(* IEC 61131-3 sources: IEC61131-3_ST_SCL_Mutation_Generator/Tests/mutatedCodeTraffic (part 2) *)

(* ---- M133.st ---- *)
FUNCTION_BLOCK TRAFFIC_CTRL

VAR_INPUT
    PedestrianButton1 : BOOL;
    PedestrianButton2 : BOOL;
END_VAR

VAR_OUTPUT
    NorthSouthRed : BOOL;
    NorthSouthYellow : BOOL;
    NorthSouthGreen : BOOL;
    EastWestRed : BOOL;
    EastWestYellow : BOOL;
    EastWestGreen : BOOL;
    PedestrianLight1 : BOOL;
    PedestrianLight2 : BOOL;
END_VAR

VAR
    LightState : INT := 0; (* 0: North-South Green, 1: North-South Yellow, 2: East-West Green, 3: East-West Yellow *)
    PedestrianRequest1 : BOOL := FALSE;
    PedestrianRequest2 : BOOL := FALSE;
    PedestrianCrossing : BOOL := FALSE;
    Timer : TON;
END_VAR

(* Check for pedestrian requests *)
IF PedestrianButton1 THEN
    PedestrianRequest1 := TRUE;
END_IF;

IF PedestrianButton2 THEN
    PedestrianRequest2 := TRUE;
END_IF;

(* Traffic light state machine *)
CASE LightState OF
    0: (* North-South Green *)
        NorthSouthGreen := TRUE;
        EastWestRed := TRUE;
        IF PedestrianRequest1 OR PedestrianRequest2 THEN
            Timer(IN := TRUE, PT := T#2s); (* Pedestrian crossing grace period *)
            IF Timer.Q THEN
                Timer(IN := FALSE);
                LightState := 2; (* MUTATED: CONST_VALUE_REPLACE *)
            END_IF;
        END_IF;

    1: (* North-South Yellow *)
        NorthSouthYellow := TRUE;
        EastWestRed := TRUE;
        Timer(IN := TRUE, PT := T#2s); (* Yellow light duration *)
        IF Timer.Q THEN
            Timer(IN := FALSE);
            LightState := 2;
        END_IF;

    2: (* East-West Green *)
        EastWestGreen := TRUE;
        NorthSouthRed := TRUE;
        IF PedestrianRequest1 THEN
            PedestrianLight1 := TRUE;
            PedestrianCrossing := TRUE;
        END_IF;
        IF PedestrianRequest2 THEN
            PedestrianLight2 := TRUE;
            PedestrianCrossing := TRUE;
        END_IF;
        IF PedestrianCrossing THEN
            Timer(IN := TRUE, PT := T#2s); (* Pedestrian crossing period *)
            IF Timer.Q THEN
                Timer(IN := FALSE);
                PedestrianRequest1 := FALSE;
                PedestrianRequest2 := FALSE;
                PedestrianLight1 := FALSE;
                PedestrianLight2 := FALSE;
                PedestrianCrossing := FALSE;
                LightState := 3;
            END_IF;
        END_IF;

    3: (* East-West Yellow *)
        EastWestYellow := TRUE;
        NorthSouthRed := TRUE;
        Timer(IN := TRUE, PT := T#2s); (* Yellow light duration *)
        IF Timer.Q THEN
            Timer(IN := FALSE);
            LightState := 0;
        END_IF;

END_CASE;

END_FUNCTION_BLOCK

(* ---- M134.st ---- *)
FUNCTION_BLOCK TRAFFIC_CTRL

VAR_INPUT
    PedestrianButton1 : BOOL;
    PedestrianButton2 : BOOL;
END_VAR

VAR_OUTPUT
    NorthSouthRed : BOOL;
    NorthSouthYellow : BOOL;
    NorthSouthGreen : BOOL;
    EastWestRed : BOOL;
    EastWestYellow : BOOL;
    EastWestGreen : BOOL;
    PedestrianLight1 : BOOL;
    PedestrianLight2 : BOOL;
END_VAR

VAR
    LightState : INT := 0; (* 0: North-South Green, 1: North-South Yellow, 2: East-West Green, 3: East-West Yellow *)
    PedestrianRequest1 : BOOL := FALSE;
    PedestrianRequest2 : BOOL := FALSE;
    PedestrianCrossing : BOOL := FALSE;
    Timer : TON;
END_VAR

(* Check for pedestrian requests *)
IF PedestrianButton1 THEN
    PedestrianRequest1 := TRUE;
END_IF;

IF PedestrianButton2 THEN
    PedestrianRequest2 := TRUE;
END_IF;

(* Traffic light state machine *)
CASE LightState OF
    0: (* North-South Green *)
        NorthSouthGreen := TRUE;
        EastWestRed := TRUE;
        IF PedestrianRequest1 OR PedestrianRequest2 THEN
            Timer(IN := TRUE, PT := T#2s); (* Pedestrian crossing grace period *)
            IF Timer.Q THEN
                Timer(IN := FALSE);
                LightState := 1;
            END_IF;
        END_IF;

    2: (* North-South Yellow *) (* MUTATED: CONST_VALUE_REPLACE *)
        NorthSouthYellow := TRUE;
        EastWestRed := TRUE;
        Timer(IN := TRUE, PT := T#2s); (* Yellow light duration *)
        IF Timer.Q THEN
            Timer(IN := FALSE);
            LightState := 2;
        END_IF;

    2: (* East-West Green *)
        EastWestGreen := TRUE;
        NorthSouthRed := TRUE;
        IF PedestrianRequest1 THEN
            PedestrianLight1 := TRUE;
            PedestrianCrossing := TRUE;
        END_IF;
        IF PedestrianRequest2 THEN
            PedestrianLight2 := TRUE;
            PedestrianCrossing := TRUE;
        END_IF;
        IF PedestrianCrossing THEN
            Timer(IN := TRUE, PT := T#2s); (* Pedestrian crossing period *)
            IF Timer.Q THEN
                Timer(IN := FALSE);
                PedestrianRequest1 := FALSE;
                PedestrianRequest2 := FALSE;
                PedestrianLight1 := FALSE;
                PedestrianLight2 := FALSE;
                PedestrianCrossing := FALSE;
                LightState := 3;
            END_IF;
        END_IF;

    3: (* East-West Yellow *)
        EastWestYellow := TRUE;
        NorthSouthRed := TRUE;
        Timer(IN := TRUE, PT := T#2s); (* Yellow light duration *)
        IF Timer.Q THEN
            Timer(IN := FALSE);
            LightState := 0;
        END_IF;

END_CASE;

END_FUNCTION_BLOCK

(* ---- M135.st ---- *)
FUNCTION_BLOCK TRAFFIC_CTRL

VAR_INPUT
    PedestrianButton1 : BOOL;
    PedestrianButton2 : BOOL;
END_VAR

VAR_OUTPUT
    NorthSouthRed : BOOL;
    NorthSouthYellow : BOOL;
    NorthSouthGreen : BOOL;
    EastWestRed : BOOL;
    EastWestYellow : BOOL;
    EastWestGreen : BOOL;
    PedestrianLight1 : BOOL;
    PedestrianLight2 : BOOL;
END_VAR

VAR
    LightState : INT := 0; (* 0: North-South Green, 1: North-South Yellow, 2: East-West Green, 3: East-West Yellow *)
    PedestrianRequest1 : BOOL := FALSE;
    PedestrianRequest2 : BOOL := FALSE;
    PedestrianCrossing : BOOL := FALSE;
    Timer : TON;
END_VAR

(* Check for pedestrian requests *)
IF PedestrianButton1 THEN
    PedestrianRequest1 := TRUE;
END_IF;

IF PedestrianButton2 THEN
    PedestrianRequest2 := TRUE;
END_IF;

(* Traffic light state machine *)
CASE LightState OF
    0: (* North-South Green *)
        NorthSouthGreen := TRUE;
        EastWestRed := TRUE;
        IF PedestrianRequest1 OR PedestrianRequest2 THEN
            Timer(IN := TRUE, PT := T#2s); (* Pedestrian crossing grace period *)
            IF Timer.Q THEN
                Timer(IN := FALSE);
                LightState := 1;
            END_IF;
        END_IF;

    1: (* North-South Yellow *)
        NorthSouthYellow := TRUE;
        EastWestRed := TRUE;
        Timer(IN := TRUE, PT := T#2s); (* Yellow light duration *)
        IF Timer.Q THEN
            Timer(IN := FALSE);
            LightState := 3; (* MUTATED: CONST_VALUE_REPLACE *)
        END_IF;

    2: (* East-West Green *)
        EastWestGreen := TRUE;
        NorthSouthRed := TRUE;
        IF PedestrianRequest1 THEN
            PedestrianLight1 := TRUE;
            PedestrianCrossing := TRUE;
        END_IF;
        IF PedestrianRequest2 THEN
            PedestrianLight2 := TRUE;
            PedestrianCrossing := TRUE;
        END_IF;
        IF PedestrianCrossing THEN
            Timer(IN := TRUE, PT := T#2s); (* Pedestrian crossing period *)
            IF Timer.Q THEN
                Timer(IN := FALSE);
                PedestrianRequest1 := FALSE;
                PedestrianRequest2 := FALSE;
                PedestrianLight1 := FALSE;
                PedestrianLight2 := FALSE;
                PedestrianCrossing := FALSE;
                LightState := 3;
            END_IF;
        END_IF;

    3: (* East-West Yellow *)
        EastWestYellow := TRUE;
        NorthSouthRed := TRUE;
        Timer(IN := TRUE, PT := T#2s); (* Yellow light duration *)
        IF Timer.Q THEN
            Timer(IN := FALSE);
            LightState := 0;
        END_IF;

END_CASE;

END_FUNCTION_BLOCK

(* ---- M136.st ---- *)
FUNCTION_BLOCK TRAFFIC_CTRL

VAR_INPUT
    PedestrianButton1 : BOOL;
    PedestrianButton2 : BOOL;
END_VAR

VAR_OUTPUT
    NorthSouthRed : BOOL;
    NorthSouthYellow : BOOL;
    NorthSouthGreen : BOOL;
    EastWestRed : BOOL;
    EastWestYellow : BOOL;
    EastWestGreen : BOOL;
    PedestrianLight1 : BOOL;
    PedestrianLight2 : BOOL;
END_VAR

VAR
    LightState : INT := 0; (* 0: North-South Green, 1: North-South Yellow, 2: East-West Green, 3: East-West Yellow *)
    PedestrianRequest1 : BOOL := FALSE;
    PedestrianRequest2 : BOOL := FALSE;
    PedestrianCrossing : BOOL := FALSE;
    Timer : TON;
END_VAR

(* Check for pedestrian requests *)
IF PedestrianButton1 THEN
    PedestrianRequest1 := TRUE;
END_IF;

IF PedestrianButton2 THEN
    PedestrianRequest2 := TRUE;
END_IF;

(* Traffic light state machine *)
CASE LightState OF
    0: (* North-South Green *)
        NorthSouthGreen := TRUE;
        EastWestRed := TRUE;
        IF PedestrianRequest1 OR PedestrianRequest2 THEN
            Timer(IN := TRUE, PT := T#2s); (* Pedestrian crossing grace period *)
            IF Timer.Q THEN
                Timer(IN := FALSE);
                LightState := 1;
            END_IF;
        END_IF;

    1: (* North-South Yellow *)
        NorthSouthYellow := TRUE;
        EastWestRed := TRUE;
        Timer(IN := TRUE, PT := T#2s); (* Yellow light duration *)
        IF Timer.Q THEN
            Timer(IN := FALSE);
            LightState := 2;
        END_IF;

    3: (* East-West Green *) (* MUTATED: CONST_VALUE_REPLACE *)
        EastWestGreen := TRUE;
        NorthSouthRed := TRUE;
        IF PedestrianRequest1 THEN
            PedestrianLight1 := TRUE;
            PedestrianCrossing := TRUE;
        END_IF;
        IF PedestrianRequest2 THEN
            PedestrianLight2 := TRUE;
            PedestrianCrossing := TRUE;
        END_IF;
        IF PedestrianCrossing THEN
            Timer(IN := TRUE, PT := T#2s); (* Pedestrian crossing period *)
            IF Timer.Q THEN
                Timer(IN := FALSE);
                PedestrianRequest1 := FALSE;
                PedestrianRequest2 := FALSE;
                PedestrianLight1 := FALSE;
                PedestrianLight2 := FALSE;
                PedestrianCrossing := FALSE;
                LightState := 3;
            END_IF;
        END_IF;

    3: (* East-West Yellow *)
        EastWestYellow := TRUE;
        NorthSouthRed := TRUE;
        Timer(IN := TRUE, PT := T#2s); (* Yellow light duration *)
        IF Timer.Q THEN
            Timer(IN := FALSE);
            LightState := 0;
        END_IF;

END_CASE;

END_FUNCTION_BLOCK

(* ---- M137.st ---- *)
FUNCTION_BLOCK TRAFFIC_CTRL

VAR_INPUT
    PedestrianButton1 : BOOL;
    PedestrianButton2 : BOOL;
END_VAR

VAR_OUTPUT
    NorthSouthRed : BOOL;
    NorthSouthYellow : BOOL;
    NorthSouthGreen : BOOL;
    EastWestRed : BOOL;
    EastWestYellow : BOOL;
    EastWestGreen : BOOL;
    PedestrianLight1 : BOOL;
    PedestrianLight2 : BOOL;
END_VAR

VAR
    LightState : INT := 0; (* 0: North-South Green, 1: North-South Yellow, 2: East-West Green, 3: East-West Yellow *)
    PedestrianRequest1 : BOOL := FALSE;
    PedestrianRequest2 : BOOL := FALSE;
    PedestrianCrossing : BOOL := FALSE;
    Timer : TON;
END_VAR

(* Check for pedestrian requests *)
IF PedestrianButton1 THEN
    PedestrianRequest1 := TRUE;
END_IF;

IF PedestrianButton2 THEN
    PedestrianRequest2 := TRUE;
END_IF;

(* Traffic light state machine *)
CASE LightState OF
    0: (* North-South Green *)
        NorthSouthGreen := TRUE;
        EastWestRed := TRUE;
        IF PedestrianRequest1 OR PedestrianRequest2 THEN
            Timer(IN := TRUE, PT := T#2s); (* Pedestrian crossing grace period *)
            IF Timer.Q THEN
                Timer(IN := FALSE);
                LightState := 1;
            END_IF;
        END_IF;

    1: (* North-South Yellow *)
        NorthSouthYellow := TRUE;
        EastWestRed := TRUE;
        Timer(IN := TRUE, PT := T#2s); (* Yellow light duration *)
        IF Timer.Q THEN
            Timer(IN := FALSE);
            LightState := 2;
        END_IF;

    2: (* East-West Green *)
        EastWestGreen := TRUE;
        NorthSouthRed := TRUE;
        IF PedestrianRequest1 THEN
            PedestrianLight1 := TRUE;
            PedestrianCrossing := TRUE;
        END_IF;
        IF PedestrianRequest2 THEN
            PedestrianLight2 := TRUE;
            PedestrianCrossing := TRUE;
        END_IF;
        IF PedestrianCrossing THEN
            Timer(IN := TRUE, PT := T#2s); (* Pedestrian crossing period *)
            IF Timer.Q THEN
                Timer(IN := FALSE);
                PedestrianRequest1 := FALSE;
                PedestrianRequest2 := FALSE;
                PedestrianLight1 := FALSE;
                PedestrianLight2 := FALSE;
                PedestrianCrossing := FALSE;
                LightState := 4; (* MUTATED: CONST_VALUE_REPLACE *)
            END_IF;
        END_IF;

    3: (* East-West Yellow *)
        EastWestYellow := TRUE;
        NorthSouthRed := TRUE;
        Timer(IN := TRUE, PT := T#2s); (* Yellow light duration *)
        IF Timer.Q THEN
            Timer(IN := FALSE);
            LightState := 0;
        END_IF;

END_CASE;

END_FUNCTION_BLOCK

(* ---- M138.st ---- *)
FUNCTION_BLOCK TRAFFIC_CTRL

VAR_INPUT
    PedestrianButton1 : BOOL;
    PedestrianButton2 : BOOL;
END_VAR

VAR_OUTPUT
    NorthSouthRed : BOOL;
    NorthSouthYellow : BOOL;
    NorthSouthGreen : BOOL;
    EastWestRed : BOOL;
    EastWestYellow : BOOL;
    EastWestGreen : BOOL;
    PedestrianLight1 : BOOL;
    PedestrianLight2 : BOOL;
END_VAR

VAR
    LightState : INT := 0; (* 0: North-South Green, 1: North-South Yellow, 2: East-West Green, 3: East-West Yellow *)
    PedestrianRequest1 : BOOL := FALSE;
    PedestrianRequest2 : BOOL := FALSE;
    PedestrianCrossing : BOOL := FALSE;
    Timer : TON;
END_VAR

(* Check for pedestrian requests *)
IF PedestrianButton1 THEN
    PedestrianRequest1 := TRUE;
END_IF;

IF PedestrianButton2 THEN
    PedestrianRequest2 := TRUE;
END_IF;

(* Traffic light state machine *)
CASE LightState OF
    0: (* North-South Green *)
        NorthSouthGreen := TRUE;
        EastWestRed := TRUE;
        IF PedestrianRequest1 OR PedestrianRequest2 THEN
            Timer(IN := TRUE, PT := T#2s); (* Pedestrian crossing grace period *)
            IF Timer.Q THEN
                Timer(IN := FALSE);
                LightState := 1;
            END_IF;
        END_IF;

    1: (* North-South Yellow *)
        NorthSouthYellow := TRUE;
        EastWestRed := TRUE;
        Timer(IN := TRUE, PT := T#2s); (* Yellow light duration *)
        IF Timer.Q THEN
            Timer(IN := FALSE);
            LightState := 2;
        END_IF;

    2: (* East-West Green *)
        EastWestGreen := TRUE;
        NorthSouthRed := TRUE;
        IF PedestrianRequest1 THEN
            PedestrianLight1 := TRUE;
            PedestrianCrossing := TRUE;
        END_IF;
        IF PedestrianRequest2 THEN
            PedestrianLight2 := TRUE;
            PedestrianCrossing := TRUE;
        END_IF;
        IF PedestrianCrossing THEN
            Timer(IN := TRUE, PT := T#2s); (* Pedestrian crossing period *)
            IF Timer.Q THEN
                Timer(IN := FALSE);
                PedestrianRequest1 := FALSE;
                PedestrianRequest2 := FALSE;
                PedestrianLight1 := FALSE;
                PedestrianLight2 := FALSE;
                PedestrianCrossing := FALSE;
                LightState := 3;
            END_IF;
        END_IF;

    4: (* East-West Yellow *) (* MUTATED: CONST_VALUE_REPLACE *)
        EastWestYellow := TRUE;
        NorthSouthRed := TRUE;
        Timer(IN := TRUE, PT := T#2s); (* Yellow light duration *)
        IF Timer.Q THEN
            Timer(IN := FALSE);
            LightState := 0;
        END_IF;

END_CASE;

END_FUNCTION_BLOCK

(* ---- M139.st ---- *)
FUNCTION_BLOCK TRAFFIC_CTRL

VAR_INPUT
    PedestrianButton1 : BOOL;
    PedestrianButton2 : BOOL;
END_VAR

VAR_OUTPUT
    NorthSouthRed : BOOL;
    NorthSouthYellow : BOOL;
    NorthSouthGreen : BOOL;
    EastWestRed : BOOL;
    EastWestYellow : BOOL;
    EastWestGreen : BOOL;
    PedestrianLight1 : BOOL;
    PedestrianLight2 : BOOL;
END_VAR

VAR
    LightState : INT := 0; (* 0: North-South Green, 1: North-South Yellow, 2: East-West Green, 3: East-West Yellow *)
    PedestrianRequest1 : BOOL := FALSE;
    PedestrianRequest2 : BOOL := FALSE;
    PedestrianCrossing : BOOL := FALSE;
    Timer : TON;
END_VAR

(* Check for pedestrian requests *)
IF PedestrianButton1 THEN
    PedestrianRequest1 := TRUE;
END_IF;

IF PedestrianButton2 THEN
    PedestrianRequest2 := TRUE;
END_IF;

(* Traffic light state machine *)
CASE LightState OF
    0: (* North-South Green *)
        NorthSouthGreen := TRUE;
        EastWestRed := TRUE;
        IF PedestrianRequest1 OR PedestrianRequest2 THEN
            Timer(IN := TRUE, PT := T#2s); (* Pedestrian crossing grace period *)
            IF Timer.Q THEN
                Timer(IN := FALSE);
                LightState := 1;
            END_IF;
        END_IF;

    1: (* North-South Yellow *)
        NorthSouthYellow := TRUE;
        EastWestRed := TRUE;
        Timer(IN := TRUE, PT := T#2s); (* Yellow light duration *)
        IF Timer.Q THEN
            Timer(IN := FALSE);
            LightState := 2;
        END_IF;

    2: (* East-West Green *)
        EastWestGreen := TRUE;
        NorthSouthRed := TRUE;
        IF PedestrianRequest1 THEN
            PedestrianLight1 := TRUE;
            PedestrianCrossing := TRUE;
        END_IF;
        IF PedestrianRequest2 THEN
            PedestrianLight2 := TRUE;
            PedestrianCrossing := TRUE;
        END_IF;
        IF PedestrianCrossing THEN
            Timer(IN := TRUE, PT := T#2s); (* Pedestrian crossing period *)
            IF Timer.Q THEN
                Timer(IN := FALSE);
                PedestrianRequest1 := FALSE;
                PedestrianRequest2 := FALSE;
                PedestrianLight1 := FALSE;
                PedestrianLight2 := FALSE;
                PedestrianCrossing := FALSE;
                LightState := 3;
            END_IF;
        END_IF;

    3: (* East-West Yellow *)
        EastWestYellow := TRUE;
        NorthSouthRed := TRUE;
        Timer(IN := TRUE, PT := T#2s); (* Yellow light duration *)
        IF Timer.Q THEN
            Timer(IN := FALSE);
            LightState := 1; (* MUTATED: CONST_VALUE_REPLACE *)
        END_IF;

END_CASE;

END_FUNCTION_BLOCK

(* ---- M140.st ---- *)
FUNCTION_BLOCK TRAFFIC_CTRL

VAR_INPUT
    PedestrianButton1 : BOOL;
    PedestrianButton2 : BOOL;
END_VAR

VAR_OUTPUT
    NorthSouthRed : BOOL;
    NorthSouthYellow : BOOL;
    NorthSouthGreen : BOOL;
    EastWestRed : BOOL;
    EastWestYellow : BOOL;
    EastWestGreen : BOOL;
    PedestrianLight1 : BOOL;
    PedestrianLight2 : BOOL;
END_VAR

VAR
    LightState : INT := 0; (* 0: North-South Green, 1: North-South Yellow, 2: East-West Green, 3: East-West Yellow *)
    PedestrianRequest1 : BOOL := FALSE;
    PedestrianRequest2 : BOOL := FALSE;
    PedestrianCrossing : BOOL := FALSE;
    Timer : TON;
END_VAR

(* Check for pedestrian requests *)
IF PedestrianButton2 THEN (* MUTATED: VAR_REPLACE *)
    PedestrianRequest1 := TRUE;
END_IF;

IF PedestrianButton2 THEN
    PedestrianRequest2 := TRUE;
END_IF;

(* Traffic light state machine *)
CASE LightState OF
    0: (* North-South Green *)
        NorthSouthGreen := TRUE;
        EastWestRed := TRUE;
        IF PedestrianRequest1 OR PedestrianRequest2 THEN
            Timer(IN := TRUE, PT := T#2s); (* Pedestrian crossing grace period *)
            IF Timer.Q THEN
                Timer(IN := FALSE);
                LightState := 1;
            END_IF;
        END_IF;

    1: (* North-South Yellow *)
        NorthSouthYellow := TRUE;
        EastWestRed := TRUE;
        Timer(IN := TRUE, PT := T#2s); (* Yellow light duration *)
        IF Timer.Q THEN
            Timer(IN := FALSE);
            LightState := 2;
        END_IF;

    2: (* East-West Green *)
        EastWestGreen := TRUE;
        NorthSouthRed := TRUE;
        IF PedestrianRequest1 THEN
            PedestrianLight1 := TRUE;
            PedestrianCrossing := TRUE;
        END_IF;
        IF PedestrianRequest2 THEN
            PedestrianLight2 := TRUE;
            PedestrianCrossing := TRUE;
        END_IF;
        IF PedestrianCrossing THEN
            Timer(IN := TRUE, PT := T#2s); (* Pedestrian crossing period *)
            IF Timer.Q THEN
                Timer(IN := FALSE);
                PedestrianRequest1 := FALSE;
                PedestrianRequest2 := FALSE;
                PedestrianLight1 := FALSE;
                PedestrianLight2 := FALSE;
                PedestrianCrossing := FALSE;
                LightState := 3;
            END_IF;
        END_IF;

    3: (* East-West Yellow *)
        EastWestYellow := TRUE;
        NorthSouthRed := TRUE;
        Timer(IN := TRUE, PT := T#2s); (* Yellow light duration *)
        IF Timer.Q THEN
            Timer(IN := FALSE);
            LightState := 0;
        END_IF;

END_CASE;

END_FUNCTION_BLOCK

(* ---- M141.st ---- *)
FUNCTION_BLOCK TRAFFIC_CTRL

VAR_INPUT
    PedestrianButton1 : BOOL;
    PedestrianButton2 : BOOL;
END_VAR

VAR_OUTPUT
    NorthSouthRed : BOOL;
    NorthSouthYellow : BOOL;
    NorthSouthGreen : BOOL;
    EastWestRed : BOOL;
    EastWestYellow : BOOL;
    EastWestGreen : BOOL;
    PedestrianLight1 : BOOL;
    PedestrianLight2 : BOOL;
END_VAR

VAR
    LightState : INT := 0; (* 0: North-South Green, 1: North-South Yellow, 2: East-West Green, 3: East-West Yellow *)
    PedestrianRequest1 : BOOL := FALSE;
    PedestrianRequest2 : BOOL := FALSE;
    PedestrianCrossing : BOOL := FALSE;
    Timer : TON;
END_VAR

(* Check for pedestrian requests *)
IF PedestrianButton1 THEN
    PedestrianRequest1 := TRUE;
END_IF;

IF NorthSouthRed THEN (* MUTATED: VAR_REPLACE *)
    PedestrianRequest2 := TRUE;
END_IF;

(* Traffic light state machine *)
CASE LightState OF
    0: (* North-South Green *)
        NorthSouthGreen := TRUE;
        EastWestRed := TRUE;
        IF PedestrianRequest1 OR PedestrianRequest2 THEN
            Timer(IN := TRUE, PT := T#2s); (* Pedestrian crossing grace period *)
            IF Timer.Q THEN
                Timer(IN := FALSE);
                LightState := 1;
            END_IF;
        END_IF;

    1: (* North-South Yellow *)
        NorthSouthYellow := TRUE;
        EastWestRed := TRUE;
        Timer(IN := TRUE, PT := T#2s); (* Yellow light duration *)
        IF Timer.Q THEN
            Timer(IN := FALSE);
            LightState := 2;
        END_IF;

    2: (* East-West Green *)
        EastWestGreen := TRUE;
        NorthSouthRed := TRUE;
        IF PedestrianRequest1 THEN
            PedestrianLight1 := TRUE;
            PedestrianCrossing := TRUE;
        END_IF;
        IF PedestrianRequest2 THEN
            PedestrianLight2 := TRUE;
            PedestrianCrossing := TRUE;
        END_IF;
        IF PedestrianCrossing THEN
            Timer(IN := TRUE, PT := T#2s); (* Pedestrian crossing period *)
            IF Timer.Q THEN
                Timer(IN := FALSE);
                PedestrianRequest1 := FALSE;
                PedestrianRequest2 := FALSE;
                PedestrianLight1 := FALSE;
                PedestrianLight2 := FALSE;
                PedestrianCrossing := FALSE;
                LightState := 3;
            END_IF;
        END_IF;

    3: (* East-West Yellow *)
        EastWestYellow := TRUE;
        NorthSouthRed := TRUE;
        Timer(IN := TRUE, PT := T#2s); (* Yellow light duration *)
        IF Timer.Q THEN
            Timer(IN := FALSE);
            LightState := 0;
        END_IF;

END_CASE;

END_FUNCTION_BLOCK

(* ---- M142.st ---- *)
FUNCTION_BLOCK TRAFFIC_CTRL

VAR_INPUT
    PedestrianButton1 : BOOL;
    PedestrianButton2 : BOOL;
END_VAR

VAR_OUTPUT
    NorthSouthRed : BOOL;
    NorthSouthYellow : BOOL;
    NorthSouthGreen : BOOL;
    EastWestRed : BOOL;
    EastWestYellow : BOOL;
    EastWestGreen : BOOL;
    PedestrianLight1 : BOOL;
    PedestrianLight2 : BOOL;
END_VAR

VAR
    LightState : INT := 0; (* 0: North-South Green, 1: North-South Yellow, 2: East-West Green, 3: East-West Yellow *)
    PedestrianRequest1 : BOOL := FALSE;
    PedestrianRequest2 : BOOL := FALSE;
    PedestrianCrossing : BOOL := FALSE;
    Timer : TON;
END_VAR

(* Check for pedestrian requests *)
IF PedestrianButton1 THEN
    PedestrianRequest1 := TRUE;
END_IF;

IF PedestrianButton2 THEN
    PedestrianRequest2 := TRUE;
END_IF;

(* Traffic light state machine *)
CASE LightState OF
    0: (* North-South Green *)
        NorthSouthGreen := TRUE;
        EastWestRed := TRUE;
        IF PedestrianRequest1 OR PedestrianRequest2 THEN
            Timer(IN := TRUE, PT := T#2s); (* Pedestrian crossing grace period *)
            IF Timer.Q THEN
                Timer(IN := FALSE);
                LightState := 1;
            END_IF;
        END_IF;

    1: (* North-South Yellow *)
        NorthSouthYellow := TRUE;
        EastWestRed := TRUE;
        Timer(IN := TRUE, PT := T#2s); (* Yellow light duration *)
        IF Timer.Q THEN
            Timer(IN := FALSE);
            LightState := 2;
        END_IF;

    2: (* East-West Green *)
        EastWestGreen := TRUE;
        NorthSouthYellow := TRUE; (* MUTATED: VAR_REPLACE *)
        IF PedestrianRequest1 THEN
            PedestrianLight1 := TRUE;
            PedestrianCrossing := TRUE;
        END_IF;
        IF PedestrianRequest2 THEN
            PedestrianLight2 := TRUE;
            PedestrianCrossing := TRUE;
        END_IF;
        IF PedestrianCrossing THEN
            Timer(IN := TRUE, PT := T#2s); (* Pedestrian crossing period *)
            IF Timer.Q THEN
                Timer(IN := FALSE);
                PedestrianRequest1 := FALSE;
                PedestrianRequest2 := FALSE;
                PedestrianLight1 := FALSE;
                PedestrianLight2 := FALSE;
                PedestrianCrossing := FALSE;
                LightState := 3;
            END_IF;
        END_IF;

    3: (* East-West Yellow *)
        EastWestYellow := TRUE;
        NorthSouthRed := TRUE;
        Timer(IN := TRUE, PT := T#2s); (* Yellow light duration *)
        IF Timer.Q THEN
            Timer(IN := FALSE);
            LightState := 0;
        END_IF;

END_CASE;

END_FUNCTION_BLOCK

(* ---- M143.st ---- *)
FUNCTION_BLOCK TRAFFIC_CTRL

VAR_INPUT
    PedestrianButton1 : BOOL;
    PedestrianButton2 : BOOL;
END_VAR

VAR_OUTPUT
    NorthSouthRed : BOOL;
    NorthSouthYellow : BOOL;
    NorthSouthGreen : BOOL;
    EastWestRed : BOOL;
    EastWestYellow : BOOL;
    EastWestGreen : BOOL;
    PedestrianLight1 : BOOL;
    PedestrianLight2 : BOOL;
END_VAR

VAR
    LightState : INT := 0; (* 0: North-South Green, 1: North-South Yellow, 2: East-West Green, 3: East-West Yellow *)
    PedestrianRequest1 : BOOL := FALSE;
    PedestrianRequest2 : BOOL := FALSE;
    PedestrianCrossing : BOOL := FALSE;
    Timer : TON;
END_VAR

(* Check for pedestrian requests *)
IF PedestrianButton1 THEN
    PedestrianRequest1 := TRUE;
END_IF;

IF PedestrianButton2 THEN
    PedestrianRequest2 := TRUE;
END_IF;

(* Traffic light state machine *)
CASE LightState OF
    0: (* North-South Green *)
        NorthSouthGreen := TRUE;
        EastWestRed := TRUE;
        IF PedestrianRequest1 OR PedestrianRequest2 THEN
            Timer(IN := TRUE, PT := T#2s); (* Pedestrian crossing grace period *)
            IF Timer.Q THEN
                Timer(IN := FALSE);
                LightState := 1;
            END_IF;
        END_IF;

    1: (* North-South Yellow *)
        NorthSouthGreen := TRUE; (* MUTATED: VAR_REPLACE *)
        EastWestRed := TRUE;
        Timer(IN := TRUE, PT := T#2s); (* Yellow light duration *)
        IF Timer.Q THEN
            Timer(IN := FALSE);
            LightState := 2;
        END_IF;

    2: (* East-West Green *)
        EastWestGreen := TRUE;
        NorthSouthRed := TRUE;
        IF PedestrianRequest1 THEN
            PedestrianLight1 := TRUE;
            PedestrianCrossing := TRUE;
        END_IF;
        IF PedestrianRequest2 THEN
            PedestrianLight2 := TRUE;
            PedestrianCrossing := TRUE;
        END_IF;
        IF PedestrianCrossing THEN
            Timer(IN := TRUE, PT := T#2s); (* Pedestrian crossing period *)
            IF Timer.Q THEN
                Timer(IN := FALSE);
                PedestrianRequest1 := FALSE;
                PedestrianRequest2 := FALSE;
                PedestrianLight1 := FALSE;
                PedestrianLight2 := FALSE;
                PedestrianCrossing := FALSE;
                LightState := 3;
            END_IF;
        END_IF;

    3: (* East-West Yellow *)
        EastWestYellow := TRUE;
        NorthSouthRed := TRUE;
        Timer(IN := TRUE, PT := T#2s); (* Yellow light duration *)
        IF Timer.Q THEN
            Timer(IN := FALSE);
            LightState := 0;
        END_IF;

END_CASE;

END_FUNCTION_BLOCK

(* ---- M144.st ---- *)
FUNCTION_BLOCK TRAFFIC_CTRL

VAR_INPUT
    PedestrianButton1 : BOOL;
    PedestrianButton2 : BOOL;
END_VAR

VAR_OUTPUT
    NorthSouthRed : BOOL;
    NorthSouthYellow : BOOL;
    NorthSouthGreen : BOOL;
    EastWestRed : BOOL;
    EastWestYellow : BOOL;
    EastWestGreen : BOOL;
    PedestrianLight1 : BOOL;
    PedestrianLight2 : BOOL;
END_VAR

VAR
    LightState : INT := 0; (* 0: North-South Green, 1: North-South Yellow, 2: East-West Green, 3: East-West Yellow *)
    PedestrianRequest1 : BOOL := FALSE;
    PedestrianRequest2 : BOOL := FALSE;
    PedestrianCrossing : BOOL := FALSE;
    Timer : TON;
END_VAR

(* Check for pedestrian requests *)
IF PedestrianButton1 THEN
    PedestrianRequest1 := TRUE;
END_IF;

IF PedestrianButton2 THEN
    PedestrianRequest2 := TRUE;
END_IF;

(* Traffic light state machine *)
CASE LightState OF
    0: (* North-South Green *)
        EastWestRed := TRUE; (* MUTATED: VAR_REPLACE *)
        EastWestRed := TRUE;
        IF PedestrianRequest1 OR PedestrianRequest2 THEN
            Timer(IN := TRUE, PT := T#2s); (* Pedestrian crossing grace period *)
            IF Timer.Q THEN
                Timer(IN := FALSE);
                LightState := 1;
            END_IF;
        END_IF;

    1: (* North-South Yellow *)
        NorthSouthYellow := TRUE;
        EastWestRed := TRUE;
        Timer(IN := TRUE, PT := T#2s); (* Yellow light duration *)
        IF Timer.Q THEN
            Timer(IN := FALSE);
            LightState := 2;
        END_IF;

    2: (* East-West Green *)
        EastWestGreen := TRUE;
        NorthSouthRed := TRUE;
        IF PedestrianRequest1 THEN
            PedestrianLight1 := TRUE;
            PedestrianCrossing := TRUE;
        END_IF;
        IF PedestrianRequest2 THEN
            PedestrianLight2 := TRUE;
            PedestrianCrossing := TRUE;
        END_IF;
        IF PedestrianCrossing THEN
            Timer(IN := TRUE, PT := T#2s); (* Pedestrian crossing period *)
            IF Timer.Q THEN
                Timer(IN := FALSE);
                PedestrianRequest1 := FALSE;
                PedestrianRequest2 := FALSE;
                PedestrianLight1 := FALSE;
                PedestrianLight2 := FALSE;
                PedestrianCrossing := FALSE;
                LightState := 3;
            END_IF;
        END_IF;

    3: (* East-West Yellow *)
        EastWestYellow := TRUE;
        NorthSouthRed := TRUE;
        Timer(IN := TRUE, PT := T#2s); (* Yellow light duration *)
        IF Timer.Q THEN
            Timer(IN := FALSE);
            LightState := 0;
        END_IF;

END_CASE;

END_FUNCTION_BLOCK

(* ---- M145.st ---- *)
FUNCTION_BLOCK TRAFFIC_CTRL

VAR_INPUT
    PedestrianButton1 : BOOL;
    PedestrianButton2 : BOOL;
END_VAR

VAR_OUTPUT
    NorthSouthRed : BOOL;
    NorthSouthYellow : BOOL;
    NorthSouthGreen : BOOL;
    EastWestRed : BOOL;
    EastWestYellow : BOOL;
    EastWestGreen : BOOL;
    PedestrianLight1 : BOOL;
    PedestrianLight2 : BOOL;
END_VAR

VAR
    LightState : INT := 0; (* 0: North-South Green, 1: North-South Yellow, 2: East-West Green, 3: East-West Yellow *)
    PedestrianRequest1 : BOOL := FALSE;
    PedestrianRequest2 : BOOL := FALSE;
    PedestrianCrossing : BOOL := FALSE;
    Timer : TON;
END_VAR

(* Check for pedestrian requests *)
IF PedestrianButton1 THEN
    PedestrianRequest1 := TRUE;
END_IF;

IF PedestrianButton2 THEN
    PedestrianRequest2 := TRUE;
END_IF;

(* Traffic light state machine *)
CASE LightState OF
    0: (* North-South Green *)
        NorthSouthGreen := TRUE;
        EastWestYellow := TRUE; (* MUTATED: VAR_REPLACE *)
        IF PedestrianRequest1 OR PedestrianRequest2 THEN
            Timer(IN := TRUE, PT := T#2s); (* Pedestrian crossing grace period *)
            IF Timer.Q THEN
                Timer(IN := FALSE);
                LightState := 1;
            END_IF;
        END_IF;

    1: (* North-South Yellow *)
        NorthSouthYellow := TRUE;
        EastWestRed := TRUE;
        Timer(IN := TRUE, PT := T#2s); (* Yellow light duration *)
        IF Timer.Q THEN
            Timer(IN := FALSE);
            LightState := 2;
        END_IF;

    2: (* East-West Green *)
        EastWestGreen := TRUE;
        NorthSouthRed := TRUE;
        IF PedestrianRequest1 THEN
            PedestrianLight1 := TRUE;
            PedestrianCrossing := TRUE;
        END_IF;
        IF PedestrianRequest2 THEN
            PedestrianLight2 := TRUE;
            PedestrianCrossing := TRUE;
        END_IF;
        IF PedestrianCrossing THEN
            Timer(IN := TRUE, PT := T#2s); (* Pedestrian crossing period *)
            IF Timer.Q THEN
                Timer(IN := FALSE);
                PedestrianRequest1 := FALSE;
                PedestrianRequest2 := FALSE;
                PedestrianLight1 := FALSE;
                PedestrianLight2 := FALSE;
                PedestrianCrossing := FALSE;
                LightState := 3;
            END_IF;
        END_IF;

    3: (* East-West Yellow *)
        EastWestYellow := TRUE;
        NorthSouthRed := TRUE;
        Timer(IN := TRUE, PT := T#2s); (* Yellow light duration *)
        IF Timer.Q THEN
            Timer(IN := FALSE);
            LightState := 0;
        END_IF;

END_CASE;

END_FUNCTION_BLOCK

(* ---- M146.st ---- *)
FUNCTION_BLOCK TRAFFIC_CTRL

VAR_INPUT
    PedestrianButton1 : BOOL;
    PedestrianButton2 : BOOL;
END_VAR

VAR_OUTPUT
    NorthSouthRed : BOOL;
    NorthSouthYellow : BOOL;
    NorthSouthGreen : BOOL;
    EastWestRed : BOOL;
    EastWestYellow : BOOL;
    EastWestGreen : BOOL;
    PedestrianLight1 : BOOL;
    PedestrianLight2 : BOOL;
END_VAR

VAR
    LightState : INT := 0; (* 0: North-South Green, 1: North-South Yellow, 2: East-West Green, 3: East-West Yellow *)
    PedestrianRequest1 : BOOL := FALSE;
    PedestrianRequest2 : BOOL := FALSE;
    PedestrianCrossing : BOOL := FALSE;
    Timer : TON;
END_VAR

(* Check for pedestrian requests *)
IF PedestrianButton1 THEN
    PedestrianRequest1 := TRUE;
END_IF;

IF PedestrianButton2 THEN
    PedestrianRequest2 := TRUE;
END_IF;

(* Traffic light state machine *)
CASE LightState OF
    0: (* North-South Green *)
        NorthSouthGreen := TRUE;
        EastWestRed := TRUE;
        IF PedestrianRequest1 OR PedestrianRequest2 THEN
            Timer(IN := TRUE, PT := T#2s); (* Pedestrian crossing grace period *)
            IF Timer.Q THEN
                Timer(IN := FALSE);
                LightState := 1;
            END_IF;
        END_IF;

    1: (* North-South Yellow *)
        NorthSouthYellow := TRUE;
        EastWestRed := TRUE;
        Timer(IN := TRUE, PT := T#2s); (* Yellow light duration *)
        IF Timer.Q THEN
            Timer(IN := FALSE);
            LightState := 2;
        END_IF;

    2: (* East-West Green *)
        EastWestGreen := TRUE;
        NorthSouthRed := TRUE;
        IF PedestrianRequest1 THEN
            PedestrianLight1 := TRUE;
            PedestrianCrossing := TRUE;
        END_IF;
        IF PedestrianRequest2 THEN
            PedestrianLight2 := TRUE;
            PedestrianCrossing := TRUE;
        END_IF;
        IF PedestrianCrossing THEN
            Timer(IN := TRUE, PT := T#2s); (* Pedestrian crossing period *)
            IF Timer.Q THEN
                Timer(IN := FALSE);
                PedestrianRequest1 := FALSE;
                PedestrianRequest2 := FALSE;
                PedestrianLight1 := FALSE;
                PedestrianLight2 := FALSE;
                PedestrianCrossing := FALSE;
                LightState := 3;
            END_IF;
        END_IF;

    3: (* East-West Yellow *)
        EastWestGreen := TRUE; (* MUTATED: VAR_REPLACE *)
        NorthSouthRed := TRUE;
        Timer(IN := TRUE, PT := T#2s); (* Yellow light duration *)
        IF Timer.Q THEN
            Timer(IN := FALSE);
            LightState := 0;
        END_IF;

END_CASE;

END_FUNCTION_BLOCK

(* ---- M147.st ---- *)
FUNCTION_BLOCK TRAFFIC_CTRL

VAR_INPUT
    PedestrianButton1 : BOOL;
    PedestrianButton2 : BOOL;
END_VAR

VAR_OUTPUT
    NorthSouthRed : BOOL;
    NorthSouthYellow : BOOL;
    NorthSouthGreen : BOOL;
    EastWestRed : BOOL;
    EastWestYellow : BOOL;
    EastWestGreen : BOOL;
    PedestrianLight1 : BOOL;
    PedestrianLight2 : BOOL;
END_VAR

VAR
    LightState : INT := 0; (* 0: North-South Green, 1: North-South Yellow, 2: East-West Green, 3: East-West Yellow *)
    PedestrianRequest1 : BOOL := FALSE;
    PedestrianRequest2 : BOOL := FALSE;
    PedestrianCrossing : BOOL := FALSE;
    Timer : TON;
END_VAR

(* Check for pedestrian requests *)
IF PedestrianButton1 THEN
    PedestrianRequest1 := TRUE;
END_IF;

IF PedestrianButton2 THEN
    PedestrianRequest2 := TRUE;
END_IF;

(* Traffic light state machine *)
CASE LightState OF
    0: (* North-South Green *)
        NorthSouthGreen := TRUE;
        EastWestRed := TRUE;
        IF PedestrianRequest1 OR PedestrianRequest2 THEN
            Timer(IN := TRUE, PT := T#2s); (* Pedestrian crossing grace period *)
            IF Timer.Q THEN
                Timer(IN := FALSE);
                LightState := 1;
            END_IF;
        END_IF;

    1: (* North-South Yellow *)
        NorthSouthYellow := TRUE;
        EastWestRed := TRUE;
        Timer(IN := TRUE, PT := T#2s); (* Yellow light duration *)
        IF Timer.Q THEN
            Timer(IN := FALSE);
            LightState := 2;
        END_IF;

    2: (* East-West Green *)
        PedestrianLight1 := TRUE; (* MUTATED: VAR_REPLACE *)
        NorthSouthRed := TRUE;
        IF PedestrianRequest1 THEN
            PedestrianLight1 := TRUE;
            PedestrianCrossing := TRUE;
        END_IF;
        IF PedestrianRequest2 THEN
            PedestrianLight2 := TRUE;
            PedestrianCrossing := TRUE;
        END_IF;
        IF PedestrianCrossing THEN
            Timer(IN := TRUE, PT := T#2s); (* Pedestrian crossing period *)
            IF Timer.Q THEN
                Timer(IN := FALSE);
                PedestrianRequest1 := FALSE;
                PedestrianRequest2 := FALSE;
                PedestrianLight1 := FALSE;
                PedestrianLight2 := FALSE;
                PedestrianCrossing := FALSE;
                LightState := 3;
            END_IF;
        END_IF;

    3: (* East-West Yellow *)
        EastWestYellow := TRUE;
        NorthSouthRed := TRUE;
        Timer(IN := TRUE, PT := T#2s); (* Yellow light duration *)
        IF Timer.Q THEN
            Timer(IN := FALSE);
            LightState := 0;
        END_IF;

END_CASE;

END_FUNCTION_BLOCK

(* ---- M148.st ---- *)
FUNCTION_BLOCK TRAFFIC_CTRL

VAR_INPUT
    PedestrianButton1 : BOOL;
    PedestrianButton2 : BOOL;
END_VAR

VAR_OUTPUT
    NorthSouthRed : BOOL;
    NorthSouthYellow : BOOL;
    NorthSouthGreen : BOOL;
    EastWestRed : BOOL;
    EastWestYellow : BOOL;
    EastWestGreen : BOOL;
    PedestrianLight1 : BOOL;
    PedestrianLight2 : BOOL;
END_VAR

VAR
    LightState : INT := 0; (* 0: North-South Green, 1: North-South Yellow, 2: East-West Green, 3: East-West Yellow *)
    PedestrianRequest1 : BOOL := FALSE;
    PedestrianRequest2 : BOOL := FALSE;
    PedestrianCrossing : BOOL := FALSE;
    Timer : TON;
END_VAR

(* Check for pedestrian requests *)
IF PedestrianButton1 THEN
    PedestrianRequest1 := TRUE;
END_IF;

IF PedestrianButton2 THEN
    PedestrianRequest2 := TRUE;
END_IF;

(* Traffic light state machine *)
CASE LightState OF
    0: (* North-South Green *)
        NorthSouthGreen := TRUE;
        EastWestRed := TRUE;
        IF PedestrianRequest1 OR PedestrianRequest2 THEN
            Timer(IN := TRUE, PT := T#2s); (* Pedestrian crossing grace period *)
            IF Timer.Q THEN
                Timer(IN := FALSE);
                LightState := 1;
            END_IF;
        END_IF;

    1: (* North-South Yellow *)
        NorthSouthYellow := TRUE;
        EastWestRed := TRUE;
        Timer(IN := TRUE, PT := T#2s); (* Yellow light duration *)
        IF Timer.Q THEN
            Timer(IN := FALSE);
            LightState := 2;
        END_IF;

    2: (* East-West Green *)
        EastWestGreen := TRUE;
        NorthSouthRed := TRUE;
        IF PedestrianRequest1 THEN
            PedestrianLight2 := TRUE; (* MUTATED: VAR_REPLACE *)
            PedestrianCrossing := TRUE;
        END_IF;
        IF PedestrianRequest2 THEN
            PedestrianLight2 := TRUE;
            PedestrianCrossing := TRUE;
        END_IF;
        IF PedestrianCrossing THEN
            Timer(IN := TRUE, PT := T#2s); (* Pedestrian crossing period *)
            IF Timer.Q THEN
                Timer(IN := FALSE);
                PedestrianRequest1 := FALSE;
                PedestrianRequest2 := FALSE;
                PedestrianLight1 := FALSE;
                PedestrianLight2 := FALSE;
                PedestrianCrossing := FALSE;
                LightState := 3;
            END_IF;
        END_IF;

    3: (* East-West Yellow *)
        EastWestYellow := TRUE;
        NorthSouthRed := TRUE;
        Timer(IN := TRUE, PT := T#2s); (* Yellow light duration *)
        IF Timer.Q THEN
            Timer(IN := FALSE);
            LightState := 0;
        END_IF;

END_CASE;

END_FUNCTION_BLOCK

(* ---- M149.st ---- *)
FUNCTION_BLOCK TRAFFIC_CTRL

VAR_INPUT
    PedestrianButton1 : BOOL;
    PedestrianButton2 : BOOL;
END_VAR

VAR_OUTPUT
    NorthSouthRed : BOOL;
    NorthSouthYellow : BOOL;
    NorthSouthGreen : BOOL;
    EastWestRed : BOOL;
    EastWestYellow : BOOL;
    EastWestGreen : BOOL;
    PedestrianLight1 : BOOL;
    PedestrianLight2 : BOOL;
END_VAR

VAR
    LightState : INT := 0; (* 0: North-South Green, 1: North-South Yellow, 2: East-West Green, 3: East-West Yellow *)
    PedestrianRequest1 : BOOL := FALSE;
    PedestrianRequest2 : BOOL := FALSE;
    PedestrianCrossing : BOOL := FALSE;
    Timer : TON;
END_VAR

(* Check for pedestrian requests *)
IF PedestrianButton1 THEN
    PedestrianRequest1 := TRUE;
END_IF;

IF PedestrianButton2 THEN
    PedestrianRequest2 := TRUE;
END_IF;

(* Traffic light state machine *)
CASE LightState OF
    0: (* North-South Green *)
        NorthSouthGreen := TRUE;
        EastWestRed := TRUE;
        IF PedestrianRequest1 OR PedestrianRequest2 THEN
            Timer(IN := TRUE, PT := T#2s); (* Pedestrian crossing grace period *)
            IF Timer.Q THEN
                Timer(IN := FALSE);
                LightState := 1;
            END_IF;
        END_IF;

    1: (* North-South Yellow *)
        NorthSouthYellow := TRUE;
        EastWestRed := TRUE;
        Timer(IN := TRUE, PT := T#2s); (* Yellow light duration *)
        IF Timer.Q THEN
            Timer(IN := FALSE);
            LightState := 2;
        END_IF;

    2: (* East-West Green *)
        EastWestGreen := TRUE;
        NorthSouthRed := TRUE;
        IF PedestrianRequest1 THEN
            PedestrianLight1 := TRUE;
            PedestrianCrossing := TRUE;
        END_IF;
        IF PedestrianRequest2 THEN
            PedestrianRequest1 := TRUE; (* MUTATED: VAR_REPLACE *)
            PedestrianCrossing := TRUE;
        END_IF;
        IF PedestrianCrossing THEN
            Timer(IN := TRUE, PT := T#2s); (* Pedestrian crossing period *)
            IF Timer.Q THEN
                Timer(IN := FALSE);
                PedestrianRequest1 := FALSE;
                PedestrianRequest2 := FALSE;
                PedestrianLight1 := FALSE;
                PedestrianLight2 := FALSE;
                PedestrianCrossing := FALSE;
                LightState := 3;
            END_IF;
        END_IF;

    3: (* East-West Yellow *)
        EastWestYellow := TRUE;
        NorthSouthRed := TRUE;
        Timer(IN := TRUE, PT := T#2s); (* Yellow light duration *)
        IF Timer.Q THEN
            Timer(IN := FALSE);
            LightState := 0;
        END_IF;

END_CASE;

END_FUNCTION_BLOCK

(* ---- M150.st ---- *)
FUNCTION_BLOCK TRAFFIC_CTRL

VAR_INPUT
    PedestrianButton1 : BOOL;
    PedestrianButton2 : BOOL;
END_VAR

VAR_OUTPUT
    NorthSouthRed : BOOL;
    NorthSouthYellow : BOOL;
    NorthSouthGreen : BOOL;
    EastWestRed : BOOL;
    EastWestYellow : BOOL;
    EastWestGreen : BOOL;
    PedestrianLight1 : BOOL;
    PedestrianLight2 : BOOL;
END_VAR

VAR
    LightState : INT := 0; (* 0: North-South Green, 1: North-South Yellow, 2: East-West Green, 3: East-West Yellow *)
    PedestrianRequest1 : BOOL := FALSE;
    PedestrianRequest2 : BOOL := FALSE;
    PedestrianCrossing : BOOL := FALSE;
    Timer : TON;
END_VAR

(* Check for pedestrian requests *)
IF PedestrianButton1 THEN
    PedestrianRequest2 := TRUE; (* MUTATED: VAR_REPLACE *)
END_IF;

IF PedestrianButton2 THEN
    PedestrianRequest2 := TRUE;
END_IF;

(* Traffic light state machine *)
CASE LightState OF
    0: (* North-South Green *)
        NorthSouthGreen := TRUE;
        EastWestRed := TRUE;
        IF PedestrianRequest1 OR PedestrianRequest2 THEN
            Timer(IN := TRUE, PT := T#2s); (* Pedestrian crossing grace period *)
            IF Timer.Q THEN
                Timer(IN := FALSE);
                LightState := 1;
            END_IF;
        END_IF;

    1: (* North-South Yellow *)
        NorthSouthYellow := TRUE;
        EastWestRed := TRUE;
        Timer(IN := TRUE, PT := T#2s); (* Yellow light duration *)
        IF Timer.Q THEN
            Timer(IN := FALSE);
            LightState := 2;
        END_IF;

    2: (* East-West Green *)
        EastWestGreen := TRUE;
        NorthSouthRed := TRUE;
        IF PedestrianRequest1 THEN
            PedestrianLight1 := TRUE;
            PedestrianCrossing := TRUE;
        END_IF;
        IF PedestrianRequest2 THEN
            PedestrianLight2 := TRUE;
            PedestrianCrossing := TRUE;
        END_IF;
        IF PedestrianCrossing THEN
            Timer(IN := TRUE, PT := T#2s); (* Pedestrian crossing period *)
            IF Timer.Q THEN
                Timer(IN := FALSE);
                PedestrianRequest1 := FALSE;
                PedestrianRequest2 := FALSE;
                PedestrianLight1 := FALSE;
                PedestrianLight2 := FALSE;
                PedestrianCrossing := FALSE;
                LightState := 3;
            END_IF;
        END_IF;

    3: (* East-West Yellow *)
        EastWestYellow := TRUE;
        NorthSouthRed := TRUE;
        Timer(IN := TRUE, PT := T#2s); (* Yellow light duration *)
        IF Timer.Q THEN
            Timer(IN := FALSE);
            LightState := 0;
        END_IF;

END_CASE;

END_FUNCTION_BLOCK

(* ---- M151.st ---- *)
FUNCTION_BLOCK TRAFFIC_CTRL

VAR_INPUT
    PedestrianButton1 : BOOL;
    PedestrianButton2 : BOOL;
END_VAR

VAR_OUTPUT
    NorthSouthRed : BOOL;
    NorthSouthYellow : BOOL;
    NorthSouthGreen : BOOL;
    EastWestRed : BOOL;
    EastWestYellow : BOOL;
    EastWestGreen : BOOL;
    PedestrianLight1 : BOOL;
    PedestrianLight2 : BOOL;
END_VAR

VAR
    LightState : INT := 0; (* 0: North-South Green, 1: North-South Yellow, 2: East-West Green, 3: East-West Yellow *)
    PedestrianRequest1 : BOOL := FALSE;
    PedestrianRequest2 : BOOL := FALSE;
    PedestrianCrossing : BOOL := FALSE;
    Timer : TON;
END_VAR

(* Check for pedestrian requests *)
IF PedestrianButton1 THEN
    PedestrianRequest1 := TRUE;
END_IF;

IF PedestrianButton2 THEN
    PedestrianCrossing := TRUE; (* MUTATED: VAR_REPLACE *)
END_IF;

(* Traffic light state machine *)
CASE LightState OF
    0: (* North-South Green *)
        NorthSouthGreen := TRUE;
        EastWestRed := TRUE;
        IF PedestrianRequest1 OR PedestrianRequest2 THEN
            Timer(IN := TRUE, PT := T#2s); (* Pedestrian crossing grace period *)
            IF Timer.Q THEN
                Timer(IN := FALSE);
                LightState := 1;
            END_IF;
        END_IF;

    1: (* North-South Yellow *)
        NorthSouthYellow := TRUE;
        EastWestRed := TRUE;
        Timer(IN := TRUE, PT := T#2s); (* Yellow light duration *)
        IF Timer.Q THEN
            Timer(IN := FALSE);
            LightState := 2;
        END_IF;

    2: (* East-West Green *)
        EastWestGreen := TRUE;
        NorthSouthRed := TRUE;
        IF PedestrianRequest1 THEN
            PedestrianLight1 := TRUE;
            PedestrianCrossing := TRUE;
        END_IF;
        IF PedestrianRequest2 THEN
            PedestrianLight2 := TRUE;
            PedestrianCrossing := TRUE;
        END_IF;
        IF PedestrianCrossing THEN
            Timer(IN := TRUE, PT := T#2s); (* Pedestrian crossing period *)
            IF Timer.Q THEN
                Timer(IN := FALSE);
                PedestrianRequest1 := FALSE;
                PedestrianRequest2 := FALSE;
                PedestrianLight1 := FALSE;
                PedestrianLight2 := FALSE;
                PedestrianCrossing := FALSE;
                LightState := 3;
            END_IF;
        END_IF;

    3: (* East-West Yellow *)
        EastWestYellow := TRUE;
        NorthSouthRed := TRUE;
        Timer(IN := TRUE, PT := T#2s); (* Yellow light duration *)
        IF Timer.Q THEN
            Timer(IN := FALSE);
            LightState := 0;
        END_IF;

END_CASE;

END_FUNCTION_BLOCK

(* ---- M152.st ---- *)
FUNCTION_BLOCK TRAFFIC_CTRL

VAR_INPUT
    PedestrianButton1 : BOOL;
    PedestrianButton2 : BOOL;
END_VAR

VAR_OUTPUT
    NorthSouthRed : BOOL;
    NorthSouthYellow : BOOL;
    NorthSouthGreen : BOOL;
    EastWestRed : BOOL;
    EastWestYellow : BOOL;
    EastWestGreen : BOOL;
    PedestrianLight1 : BOOL;
    PedestrianLight2 : BOOL;
END_VAR

VAR
    LightState : INT := 0; (* 0: North-South Green, 1: North-South Yellow, 2: East-West Green, 3: East-West Yellow *)
    PedestrianRequest1 : BOOL := FALSE;
    PedestrianRequest2 : BOOL := FALSE;
    PedestrianCrossing : BOOL := FALSE;
    Timer : TON;
END_VAR

(* Check for pedestrian requests *)
IF PedestrianButton1 THEN
    PedestrianRequest1 := TRUE;
END_IF;

IF PedestrianButton2 THEN
    PedestrianRequest2 := TRUE;
END_IF;

(* Traffic light state machine *)
CASE LightState OF
    0: (* North-South Green *)
        NorthSouthGreen := TRUE;
        EastWestRed := TRUE;
        IF PedestrianRequest1 OR PedestrianRequest2 THEN
            Timer(IN := TRUE, PT := T#2s); (* Pedestrian crossing grace period *)
            IF Timer.Q THEN
                Timer(IN := FALSE);
                LightState := 1;
            END_IF;
        END_IF;

    1: (* North-South Yellow *)
        NorthSouthYellow := TRUE;
        EastWestRed := TRUE;
        Timer(IN := TRUE, PT := T#2s); (* Yellow light duration *)
        IF Timer.Q THEN
            Timer(IN := FALSE);
            LightState := 2;
        END_IF;

    2: (* East-West Green *)
        EastWestGreen := TRUE;
        NorthSouthRed := TRUE;
        IF PedestrianRequest1 THEN
            PedestrianLight1 := TRUE;
            PedestrianButton1 := TRUE; (* MUTATED: VAR_REPLACE *)
        END_IF;
        IF PedestrianRequest2 THEN
            PedestrianLight2 := TRUE;
            PedestrianCrossing := TRUE;
        END_IF;
        IF PedestrianCrossing THEN
            Timer(IN := TRUE, PT := T#2s); (* Pedestrian crossing period *)
            IF Timer.Q THEN
                Timer(IN := FALSE);
                PedestrianRequest1 := FALSE;
                PedestrianRequest2 := FALSE;
                PedestrianLight1 := FALSE;
                PedestrianLight2 := FALSE;
                PedestrianCrossing := FALSE;
                LightState := 3;
            END_IF;
        END_IF;

    3: (* East-West Yellow *)
        EastWestYellow := TRUE;
        NorthSouthRed := TRUE;
        Timer(IN := TRUE, PT := T#2s); (* Yellow light duration *)
        IF Timer.Q THEN
            Timer(IN := FALSE);
            LightState := 0;
        END_IF;

END_CASE;

END_FUNCTION_BLOCK

(* ---- M153.st ---- *)
FUNCTION_BLOCK TRAFFIC_CTRL

VAR_INPUT
    PedestrianButton1 : BOOL;
    PedestrianButton2 : BOOL;
END_VAR

VAR_OUTPUT
    NorthSouthRed : BOOL;
    NorthSouthYellow : BOOL;
    NorthSouthGreen : BOOL;
    EastWestRed : BOOL;
    EastWestYellow : BOOL;
    EastWestGreen : BOOL;
    PedestrianLight1 : BOOL;
    PedestrianLight2 : BOOL;
END_VAR

VAR
    LightState : INT := 0; (* 0: North-South Green, 1: North-South Yellow, 2: East-West Green, 3: East-West Yellow *)
    PedestrianRequest1 : BOOL := FALSE;
    PedestrianRequest2 : BOOL := FALSE;
    PedestrianCrossing : BOOL := FALSE;
    Timer : TON;
END_VAR

(* Check for pedestrian requests *)
IF PedestrianButton1 THEN
    PedestrianRequest1 := NOT (TRUE); (* MUTATED: ASSIGN_NEGATE *)
END_IF;

IF PedestrianButton2 THEN
    PedestrianRequest2 := TRUE;
END_IF;

(* Traffic light state machine *)
CASE LightState OF
    0: (* North-South Green *)
        NorthSouthGreen := TRUE;
        EastWestRed := TRUE;
        IF PedestrianRequest1 OR PedestrianRequest2 THEN
            Timer(IN := TRUE, PT := T#2s); (* Pedestrian crossing grace period *)
            IF Timer.Q THEN
                Timer(IN := FALSE);
                LightState := 1;
            END_IF;
        END_IF;

    1: (* North-South Yellow *)
        NorthSouthYellow := TRUE;
        EastWestRed := TRUE;
        Timer(IN := TRUE, PT := T#2s); (* Yellow light duration *)
        IF Timer.Q THEN
            Timer(IN := FALSE);
            LightState := 2;
        END_IF;

    2: (* East-West Green *)
        EastWestGreen := TRUE;
        NorthSouthRed := TRUE;
        IF PedestrianRequest1 THEN
            PedestrianLight1 := TRUE;
            PedestrianCrossing := TRUE;
        END_IF;
        IF PedestrianRequest2 THEN
            PedestrianLight2 := TRUE;
            PedestrianCrossing := TRUE;
        END_IF;
        IF PedestrianCrossing THEN
            Timer(IN := TRUE, PT := T#2s); (* Pedestrian crossing period *)
            IF Timer.Q THEN
                Timer(IN := FALSE);
                PedestrianRequest1 := FALSE;
                PedestrianRequest2 := FALSE;
                PedestrianLight1 := FALSE;
                PedestrianLight2 := FALSE;
                PedestrianCrossing := FALSE;
                LightState := 3;
            END_IF;
        END_IF;

    3: (* East-West Yellow *)
        EastWestYellow := TRUE;
        NorthSouthRed := TRUE;
        Timer(IN := TRUE, PT := T#2s); (* Yellow light duration *)
        IF Timer.Q THEN
            Timer(IN := FALSE);
            LightState := 0;
        END_IF;

END_CASE;

END_FUNCTION_BLOCK

(* ---- M154.st ---- *)
FUNCTION_BLOCK TRAFFIC_CTRL

VAR_INPUT
    PedestrianButton1 : BOOL;
    PedestrianButton2 : BOOL;
END_VAR

VAR_OUTPUT
    NorthSouthRed : BOOL;
    NorthSouthYellow : BOOL;
    NorthSouthGreen : BOOL;
    EastWestRed : BOOL;
    EastWestYellow : BOOL;
    EastWestGreen : BOOL;
    PedestrianLight1 : BOOL;
    PedestrianLight2 : BOOL;
END_VAR

VAR
    LightState : INT := 0; (* 0: North-South Green, 1: North-South Yellow, 2: East-West Green, 3: East-West Yellow *)
    PedestrianRequest1 : BOOL := FALSE;
    PedestrianRequest2 : BOOL := FALSE;
    PedestrianCrossing : BOOL := FALSE;
    Timer : TON;
END_VAR

(* Check for pedestrian requests *)
IF PedestrianButton1 THEN
    PedestrianRequest1 := TRUE;
END_IF;

IF PedestrianButton2 THEN
    PedestrianRequest2 := NOT (TRUE); (* MUTATED: ASSIGN_NEGATE *)
END_IF;

(* Traffic light state machine *)
CASE LightState OF
    0: (* North-South Green *)
        NorthSouthGreen := TRUE;
        EastWestRed := TRUE;
        IF PedestrianRequest1 OR PedestrianRequest2 THEN
            Timer(IN := TRUE, PT := T#2s); (* Pedestrian crossing grace period *)
            IF Timer.Q THEN
                Timer(IN := FALSE);
                LightState := 1;
            END_IF;
        END_IF;

    1: (* North-South Yellow *)
        NorthSouthYellow := TRUE;
        EastWestRed := TRUE;
        Timer(IN := TRUE, PT := T#2s); (* Yellow light duration *)
        IF Timer.Q THEN
            Timer(IN := FALSE);
            LightState := 2;
        END_IF;

    2: (* East-West Green *)
        EastWestGreen := TRUE;
        NorthSouthRed := TRUE;
        IF PedestrianRequest1 THEN
            PedestrianLight1 := TRUE;
            PedestrianCrossing := TRUE;
        END_IF;
        IF PedestrianRequest2 THEN
            PedestrianLight2 := TRUE;
            PedestrianCrossing := TRUE;
        END_IF;
        IF PedestrianCrossing THEN
            Timer(IN := TRUE, PT := T#2s); (* Pedestrian crossing period *)
            IF Timer.Q THEN
                Timer(IN := FALSE);
                PedestrianRequest1 := FALSE;
                PedestrianRequest2 := FALSE;
                PedestrianLight1 := FALSE;
                PedestrianLight2 := FALSE;
                PedestrianCrossing := FALSE;
                LightState := 3;
            END_IF;
        END_IF;

    3: (* East-West Yellow *)
        EastWestYellow := TRUE;
        NorthSouthRed := TRUE;
        Timer(IN := TRUE, PT := T#2s); (* Yellow light duration *)
        IF Timer.Q THEN
            Timer(IN := FALSE);
            LightState := 0;
        END_IF;

END_CASE;

END_FUNCTION_BLOCK

(* ---- M155.st ---- *)
FUNCTION_BLOCK TRAFFIC_CTRL

VAR_INPUT
    PedestrianButton1 : BOOL;
    PedestrianButton2 : BOOL;
END_VAR

VAR_OUTPUT
    NorthSouthRed : BOOL;
    NorthSouthYellow : BOOL;
    NorthSouthGreen : BOOL;
    EastWestRed : BOOL;
    EastWestYellow : BOOL;
    EastWestGreen : BOOL;
    PedestrianLight1 : BOOL;
    PedestrianLight2 : BOOL;
END_VAR

VAR
    LightState : INT := 0; (* 0: North-South Green, 1: North-South Yellow, 2: East-West Green, 3: East-West Yellow *)
    PedestrianRequest1 : BOOL := FALSE;
    PedestrianRequest2 : BOOL := FALSE;
    PedestrianCrossing : BOOL := FALSE;
    Timer : TON;
END_VAR

(* Check for pedestrian requests *)
IF PedestrianButton1 THEN
    PedestrianRequest1 := TRUE;
END_IF;

IF PedestrianButton2 THEN
    PedestrianRequest2 := TRUE;
END_IF;

(* Traffic light state machine *)
CASE LightState OF
    0: (* North-South Green *)
        NorthSouthGreen := NOT (TRUE); (* MUTATED: ASSIGN_NEGATE *)
        EastWestRed := TRUE;
        IF PedestrianRequest1 OR PedestrianRequest2 THEN
            Timer(IN := TRUE, PT := T#2s); (* Pedestrian crossing grace period *)
            IF Timer.Q THEN
                Timer(IN := FALSE);
                LightState := 1;
            END_IF;
        END_IF;

    1: (* North-South Yellow *)
        NorthSouthYellow := TRUE;
        EastWestRed := TRUE;
        Timer(IN := TRUE, PT := T#2s); (* Yellow light duration *)
        IF Timer.Q THEN
            Timer(IN := FALSE);
            LightState := 2;
        END_IF;

    2: (* East-West Green *)
        EastWestGreen := TRUE;
        NorthSouthRed := TRUE;
        IF PedestrianRequest1 THEN
            PedestrianLight1 := TRUE;
            PedestrianCrossing := TRUE;
        END_IF;
        IF PedestrianRequest2 THEN
            PedestrianLight2 := TRUE;
            PedestrianCrossing := TRUE;
        END_IF;
        IF PedestrianCrossing THEN
            Timer(IN := TRUE, PT := T#2s); (* Pedestrian crossing period *)
            IF Timer.Q THEN
                Timer(IN := FALSE);
                PedestrianRequest1 := FALSE;
                PedestrianRequest2 := FALSE;
                PedestrianLight1 := FALSE;
                PedestrianLight2 := FALSE;
                PedestrianCrossing := FALSE;
                LightState := 3;
            END_IF;
        END_IF;

    3: (* East-West Yellow *)
        EastWestYellow := TRUE;
        NorthSouthRed := TRUE;
        Timer(IN := TRUE, PT := T#2s); (* Yellow light duration *)
        IF Timer.Q THEN
            Timer(IN := FALSE);
            LightState := 0;
        END_IF;

END_CASE;

END_FUNCTION_BLOCK

(* ---- M156.st ---- *)
FUNCTION_BLOCK TRAFFIC_CTRL

VAR_INPUT
    PedestrianButton1 : BOOL;
    PedestrianButton2 : BOOL;
END_VAR

VAR_OUTPUT
    NorthSouthRed : BOOL;
    NorthSouthYellow : BOOL;
    NorthSouthGreen : BOOL;
    EastWestRed : BOOL;
    EastWestYellow : BOOL;
    EastWestGreen : BOOL;
    PedestrianLight1 : BOOL;
    PedestrianLight2 : BOOL;
END_VAR

VAR
    LightState : INT := 0; (* 0: North-South Green, 1: North-South Yellow, 2: East-West Green, 3: East-West Yellow *)
    PedestrianRequest1 : BOOL := FALSE;
    PedestrianRequest2 : BOOL := FALSE;
    PedestrianCrossing : BOOL := FALSE;
    Timer : TON;
END_VAR

(* Check for pedestrian requests *)
IF PedestrianButton1 THEN
    PedestrianRequest1 := TRUE;
END_IF;

IF PedestrianButton2 THEN
    PedestrianRequest2 := TRUE;
END_IF;

(* Traffic light state machine *)
CASE LightState OF
    0: (* North-South Green *)
        NorthSouthGreen := TRUE;
        EastWestRed := NOT (TRUE); (* MUTATED: ASSIGN_NEGATE *)
        IF PedestrianRequest1 OR PedestrianRequest2 THEN
            Timer(IN := TRUE, PT := T#2s); (* Pedestrian crossing grace period *)
            IF Timer.Q THEN
                Timer(IN := FALSE);
                LightState := 1;
            END_IF;
        END_IF;

    1: (* North-South Yellow *)
        NorthSouthYellow := TRUE;
        EastWestRed := TRUE;
        Timer(IN := TRUE, PT := T#2s); (* Yellow light duration *)
        IF Timer.Q THEN
            Timer(IN := FALSE);
            LightState := 2;
        END_IF;

    2: (* East-West Green *)
        EastWestGreen := TRUE;
        NorthSouthRed := TRUE;
        IF PedestrianRequest1 THEN
            PedestrianLight1 := TRUE;
            PedestrianCrossing := TRUE;
        END_IF;
        IF PedestrianRequest2 THEN
            PedestrianLight2 := TRUE;
            PedestrianCrossing := TRUE;
        END_IF;
        IF PedestrianCrossing THEN
            Timer(IN := TRUE, PT := T#2s); (* Pedestrian crossing period *)
            IF Timer.Q THEN
                Timer(IN := FALSE);
                PedestrianRequest1 := FALSE;
                PedestrianRequest2 := FALSE;
                PedestrianLight1 := FALSE;
                PedestrianLight2 := FALSE;
                PedestrianCrossing := FALSE;
                LightState := 3;
            END_IF;
        END_IF;

    3: (* East-West Yellow *)
        EastWestYellow := TRUE;
        NorthSouthRed := TRUE;
        Timer(IN := TRUE, PT := T#2s); (* Yellow light duration *)
        IF Timer.Q THEN
            Timer(IN := FALSE);
            LightState := 0;
        END_IF;

END_CASE;

END_FUNCTION_BLOCK

(* ---- M157.st ---- *)
FUNCTION_BLOCK TRAFFIC_CTRL

VAR_INPUT
    PedestrianButton1 : BOOL;
    PedestrianButton2 : BOOL;
END_VAR

VAR_OUTPUT
    NorthSouthRed : BOOL;
    NorthSouthYellow : BOOL;
    NorthSouthGreen : BOOL;
    EastWestRed : BOOL;
    EastWestYellow : BOOL;
    EastWestGreen : BOOL;
    PedestrianLight1 : BOOL;
    PedestrianLight2 : BOOL;
END_VAR

VAR
    LightState : INT := 0; (* 0: North-South Green, 1: North-South Yellow, 2: East-West Green, 3: East-West Yellow *)
    PedestrianRequest1 : BOOL := FALSE;
    PedestrianRequest2 : BOOL := FALSE;
    PedestrianCrossing : BOOL := FALSE;
    Timer : TON;
END_VAR

(* Check for pedestrian requests *)
IF PedestrianButton1 THEN
    PedestrianRequest1 := TRUE;
END_IF;

IF PedestrianButton2 THEN
    PedestrianRequest2 := TRUE;
END_IF;

(* Traffic light state machine *)
CASE LightState OF
    0: (* North-South Green *)
        NorthSouthGreen := TRUE;
        EastWestRed := TRUE;
        IF PedestrianRequest1 OR PedestrianRequest2 THEN
            Timer(IN := TRUE, PT := T#2s); (* Pedestrian crossing grace period *)
            IF Timer.Q THEN
                Timer(IN := FALSE);
                LightState := 1;
            END_IF;
        END_IF;

    1: (* North-South Yellow *)
        NorthSouthYellow := NOT (TRUE); (* MUTATED: ASSIGN_NEGATE *)
        EastWestRed := TRUE;
        Timer(IN := TRUE, PT := T#2s); (* Yellow light duration *)
        IF Timer.Q THEN
            Timer(IN := FALSE);
            LightState := 2;
        END_IF;

    2: (* East-West Green *)
        EastWestGreen := TRUE;
        NorthSouthRed := TRUE;
        IF PedestrianRequest1 THEN
            PedestrianLight1 := TRUE;
            PedestrianCrossing := TRUE;
        END_IF;
        IF PedestrianRequest2 THEN
            PedestrianLight2 := TRUE;
            PedestrianCrossing := TRUE;
        END_IF;
        IF PedestrianCrossing THEN
            Timer(IN := TRUE, PT := T#2s); (* Pedestrian crossing period *)
            IF Timer.Q THEN
                Timer(IN := FALSE);
                PedestrianRequest1 := FALSE;
                PedestrianRequest2 := FALSE;
                PedestrianLight1 := FALSE;
                PedestrianLight2 := FALSE;
                PedestrianCrossing := FALSE;
                LightState := 3;
            END_IF;
        END_IF;

    3: (* East-West Yellow *)
        EastWestYellow := TRUE;
        NorthSouthRed := TRUE;
        Timer(IN := TRUE, PT := T#2s); (* Yellow light duration *)
        IF Timer.Q THEN
            Timer(IN := FALSE);
            LightState := 0;
        END_IF;

END_CASE;

END_FUNCTION_BLOCK

(* ---- M158.st ---- *)
FUNCTION_BLOCK TRAFFIC_CTRL

VAR_INPUT
    PedestrianButton1 : BOOL;
    PedestrianButton2 : BOOL;
END_VAR

VAR_OUTPUT
    NorthSouthRed : BOOL;
    NorthSouthYellow : BOOL;
    NorthSouthGreen : BOOL;
    EastWestRed : BOOL;
    EastWestYellow : BOOL;
    EastWestGreen : BOOL;
    PedestrianLight1 : BOOL;
    PedestrianLight2 : BOOL;
END_VAR

VAR
    LightState : INT := 0; (* 0: North-South Green, 1: North-South Yellow, 2: East-West Green, 3: East-West Yellow *)
    PedestrianRequest1 : BOOL := FALSE;
    PedestrianRequest2 : BOOL := FALSE;
    PedestrianCrossing : BOOL := FALSE;
    Timer : TON;
END_VAR

(* Check for pedestrian requests *)
IF PedestrianButton1 THEN
    PedestrianRequest1 := TRUE;
END_IF;

IF PedestrianButton2 THEN
    PedestrianRequest2 := TRUE;
END_IF;

(* Traffic light state machine *)
CASE LightState OF
    0: (* North-South Green *)
        NorthSouthGreen := TRUE;
        EastWestRed := TRUE;
        IF PedestrianRequest1 OR PedestrianRequest2 THEN
            Timer(IN := TRUE, PT := T#2s); (* Pedestrian crossing grace period *)
            IF Timer.Q THEN
                Timer(IN := FALSE);
                LightState := 1;
            END_IF;
        END_IF;

    1: (* North-South Yellow *)
        NorthSouthYellow := TRUE;
        EastWestRed := NOT (TRUE); (* MUTATED: ASSIGN_NEGATE *)
        Timer(IN := TRUE, PT := T#2s); (* Yellow light duration *)
        IF Timer.Q THEN
            Timer(IN := FALSE);
            LightState := 2;
        END_IF;

    2: (* East-West Green *)
        EastWestGreen := TRUE;
        NorthSouthRed := TRUE;
        IF PedestrianRequest1 THEN
            PedestrianLight1 := TRUE;
            PedestrianCrossing := TRUE;
        END_IF;
        IF PedestrianRequest2 THEN
            PedestrianLight2 := TRUE;
            PedestrianCrossing := TRUE;
        END_IF;
        IF PedestrianCrossing THEN
            Timer(IN := TRUE, PT := T#2s); (* Pedestrian crossing period *)
            IF Timer.Q THEN
                Timer(IN := FALSE);
                PedestrianRequest1 := FALSE;
                PedestrianRequest2 := FALSE;
                PedestrianLight1 := FALSE;
                PedestrianLight2 := FALSE;
                PedestrianCrossing := FALSE;
                LightState := 3;
            END_IF;
        END_IF;

    3: (* East-West Yellow *)
        EastWestYellow := TRUE;
        NorthSouthRed := TRUE;
        Timer(IN := TRUE, PT := T#2s); (* Yellow light duration *)
        IF Timer.Q THEN
            Timer(IN := FALSE);
            LightState := 0;
        END_IF;

END_CASE;

END_FUNCTION_BLOCK

(* ---- M159.st ---- *)
FUNCTION_BLOCK TRAFFIC_CTRL

VAR_INPUT
    PedestrianButton1 : BOOL;
    PedestrianButton2 : BOOL;
END_VAR

VAR_OUTPUT
    NorthSouthRed : BOOL;
    NorthSouthYellow : BOOL;
    NorthSouthGreen : BOOL;
    EastWestRed : BOOL;
    EastWestYellow : BOOL;
    EastWestGreen : BOOL;
    PedestrianLight1 : BOOL;
    PedestrianLight2 : BOOL;
END_VAR

VAR
    LightState : INT := 0; (* 0: North-South Green, 1: North-South Yellow, 2: East-West Green, 3: East-West Yellow *)
    PedestrianRequest1 : BOOL := FALSE;
    PedestrianRequest2 : BOOL := FALSE;
    PedestrianCrossing : BOOL := FALSE;
    Timer : TON;
END_VAR

(* Check for pedestrian requests *)
IF PedestrianButton1 THEN
    PedestrianRequest1 := TRUE;
END_IF;

IF PedestrianButton2 THEN
    PedestrianRequest2 := TRUE;
END_IF;

(* Traffic light state machine *)
CASE LightState OF
    0: (* North-South Green *)
        NorthSouthGreen := TRUE;
        EastWestRed := TRUE;
        IF PedestrianRequest1 OR PedestrianRequest2 THEN
            Timer(IN := TRUE, PT := T#2s); (* Pedestrian crossing grace period *)
            IF Timer.Q THEN
                Timer(IN := FALSE);
                LightState := 1;
            END_IF;
        END_IF;

    1: (* North-South Yellow *)
        NorthSouthYellow := TRUE;
        EastWestRed := TRUE;
        Timer(IN := TRUE, PT := T#2s); (* Yellow light duration *)
        IF Timer.Q THEN
            Timer(IN := FALSE);
            LightState := 2;
        END_IF;

    2: (* East-West Green *)
        EastWestGreen := NOT (TRUE); (* MUTATED: ASSIGN_NEGATE *)
        NorthSouthRed := TRUE;
        IF PedestrianRequest1 THEN
            PedestrianLight1 := TRUE;
            PedestrianCrossing := TRUE;
        END_IF;
        IF PedestrianRequest2 THEN
            PedestrianLight2 := TRUE;
            PedestrianCrossing := TRUE;
        END_IF;
        IF PedestrianCrossing THEN
            Timer(IN := TRUE, PT := T#2s); (* Pedestrian crossing period *)
            IF Timer.Q THEN
                Timer(IN := FALSE);
                PedestrianRequest1 := FALSE;
                PedestrianRequest2 := FALSE;
                PedestrianLight1 := FALSE;
                PedestrianLight2 := FALSE;
                PedestrianCrossing := FALSE;
                LightState := 3;
            END_IF;
        END_IF;

    3: (* East-West Yellow *)
        EastWestYellow := TRUE;
        NorthSouthRed := TRUE;
        Timer(IN := TRUE, PT := T#2s); (* Yellow light duration *)
        IF Timer.Q THEN
            Timer(IN := FALSE);
            LightState := 0;
        END_IF;

END_CASE;

END_FUNCTION_BLOCK

(* ---- M160.st ---- *)
FUNCTION_BLOCK TRAFFIC_CTRL

VAR_INPUT
    PedestrianButton1 : BOOL;
    PedestrianButton2 : BOOL;
END_VAR

VAR_OUTPUT
    NorthSouthRed : BOOL;
    NorthSouthYellow : BOOL;
    NorthSouthGreen : BOOL;
    EastWestRed : BOOL;
    EastWestYellow : BOOL;
    EastWestGreen : BOOL;
    PedestrianLight1 : BOOL;
    PedestrianLight2 : BOOL;
END_VAR

VAR
    LightState : INT := 0; (* 0: North-South Green, 1: North-South Yellow, 2: East-West Green, 3: East-West Yellow *)
    PedestrianRequest1 : BOOL := FALSE;
    PedestrianRequest2 : BOOL := FALSE;
    PedestrianCrossing : BOOL := FALSE;
    Timer : TON;
END_VAR

(* Check for pedestrian requests *)
IF PedestrianButton1 THEN
    PedestrianRequest1 := TRUE;
END_IF;

IF PedestrianButton2 THEN
    PedestrianRequest2 := TRUE;
END_IF;

(* Traffic light state machine *)
CASE LightState OF
    0: (* North-South Green *)
        NorthSouthGreen := TRUE;
        EastWestRed := TRUE;
        IF PedestrianRequest1 OR PedestrianRequest2 THEN
            Timer(IN := TRUE, PT := T#2s); (* Pedestrian crossing grace period *)
            IF Timer.Q THEN
                Timer(IN := FALSE);
                LightState := 1;
            END_IF;
        END_IF;

    1: (* North-South Yellow *)
        NorthSouthYellow := TRUE;
        EastWestRed := TRUE;
        Timer(IN := TRUE, PT := T#2s); (* Yellow light duration *)
        IF Timer.Q THEN
            Timer(IN := FALSE);
            LightState := 2;
        END_IF;

    2: (* East-West Green *)
        EastWestGreen := TRUE;
        NorthSouthRed := NOT (TRUE); (* MUTATED: ASSIGN_NEGATE *)
        IF PedestrianRequest1 THEN
            PedestrianLight1 := TRUE;
            PedestrianCrossing := TRUE;
        END_IF;
        IF PedestrianRequest2 THEN
            PedestrianLight2 := TRUE;
            PedestrianCrossing := TRUE;
        END_IF;
        IF PedestrianCrossing THEN
            Timer(IN := TRUE, PT := T#2s); (* Pedestrian crossing period *)
            IF Timer.Q THEN
                Timer(IN := FALSE);
                PedestrianRequest1 := FALSE;
                PedestrianRequest2 := FALSE;
                PedestrianLight1 := FALSE;
                PedestrianLight2 := FALSE;
                PedestrianCrossing := FALSE;
                LightState := 3;
            END_IF;
        END_IF;

    3: (* East-West Yellow *)
        EastWestYellow := TRUE;
        NorthSouthRed := TRUE;
        Timer(IN := TRUE, PT := T#2s); (* Yellow light duration *)
        IF Timer.Q THEN
            Timer(IN := FALSE);
            LightState := 0;
        END_IF;

END_CASE;

END_FUNCTION_BLOCK

(* ---- M161.st ---- *)
FUNCTION_BLOCK TRAFFIC_CTRL

VAR_INPUT
    PedestrianButton1 : BOOL;
    PedestrianButton2 : BOOL;
END_VAR

VAR_OUTPUT
    NorthSouthRed : BOOL;
    NorthSouthYellow : BOOL;
    NorthSouthGreen : BOOL;
    EastWestRed : BOOL;
    EastWestYellow : BOOL;
    EastWestGreen : BOOL;
    PedestrianLight1 : BOOL;
    PedestrianLight2 : BOOL;
END_VAR

VAR
    LightState : INT := 0; (* 0: North-South Green, 1: North-South Yellow, 2: East-West Green, 3: East-West Yellow *)
    PedestrianRequest1 : BOOL := FALSE;
    PedestrianRequest2 : BOOL := FALSE;
    PedestrianCrossing : BOOL := FALSE;
    Timer : TON;
END_VAR

(* Check for pedestrian requests *)
IF PedestrianButton1 THEN
    PedestrianRequest1 := TRUE;
END_IF;

IF PedestrianButton2 THEN
    PedestrianRequest2 := TRUE;
END_IF;

(* Traffic light state machine *)
CASE LightState OF
    0: (* North-South Green *)
        NorthSouthGreen := TRUE;
        EastWestRed := TRUE;
        IF PedestrianRequest1 OR PedestrianRequest2 THEN
            Timer(IN := TRUE, PT := T#2s); (* Pedestrian crossing grace period *)
            IF Timer.Q THEN
                Timer(IN := FALSE);
                LightState := 1;
            END_IF;
        END_IF;

    1: (* North-South Yellow *)
        NorthSouthYellow := TRUE;
        EastWestRed := TRUE;
        Timer(IN := TRUE, PT := T#2s); (* Yellow light duration *)
        IF Timer.Q THEN
            Timer(IN := FALSE);
            LightState := 2;
        END_IF;

    2: (* East-West Green *)
        EastWestGreen := TRUE;
        NorthSouthRed := TRUE;
        IF PedestrianRequest1 THEN
            PedestrianLight1 := NOT (TRUE); (* MUTATED: ASSIGN_NEGATE *)
            PedestrianCrossing := TRUE;
        END_IF;
        IF PedestrianRequest2 THEN
            PedestrianLight2 := TRUE;
            PedestrianCrossing := TRUE;
        END_IF;
        IF PedestrianCrossing THEN
            Timer(IN := TRUE, PT := T#2s); (* Pedestrian crossing period *)
            IF Timer.Q THEN
                Timer(IN := FALSE);
                PedestrianRequest1 := FALSE;
                PedestrianRequest2 := FALSE;
                PedestrianLight1 := FALSE;
                PedestrianLight2 := FALSE;
                PedestrianCrossing := FALSE;
                LightState := 3;
            END_IF;
        END_IF;

    3: (* East-West Yellow *)
        EastWestYellow := TRUE;
        NorthSouthRed := TRUE;
        Timer(IN := TRUE, PT := T#2s); (* Yellow light duration *)
        IF Timer.Q THEN
            Timer(IN := FALSE);
            LightState := 0;
        END_IF;

END_CASE;

END_FUNCTION_BLOCK

(* ---- M162.st ---- *)
FUNCTION_BLOCK TRAFFIC_CTRL

VAR_INPUT
    PedestrianButton1 : BOOL;
    PedestrianButton2 : BOOL;
END_VAR

VAR_OUTPUT
    NorthSouthRed : BOOL;
    NorthSouthYellow : BOOL;
    NorthSouthGreen : BOOL;
    EastWestRed : BOOL;
    EastWestYellow : BOOL;
    EastWestGreen : BOOL;
    PedestrianLight1 : BOOL;
    PedestrianLight2 : BOOL;
END_VAR

VAR
    LightState : INT := 0; (* 0: North-South Green, 1: North-South Yellow, 2: East-West Green, 3: East-West Yellow *)
    PedestrianRequest1 : BOOL := FALSE;
    PedestrianRequest2 : BOOL := FALSE;
    PedestrianCrossing : BOOL := FALSE;
    Timer : TON;
END_VAR

(* Check for pedestrian requests *)
IF PedestrianButton1 THEN
    PedestrianRequest1 := TRUE;
END_IF;

IF PedestrianButton2 THEN
    PedestrianRequest2 := TRUE;
END_IF;

(* Traffic light state machine *)
CASE LightState OF
    0: (* North-South Green *)
        NorthSouthGreen := TRUE;
        EastWestRed := TRUE;
        IF PedestrianRequest1 OR PedestrianRequest2 THEN
            Timer(IN := TRUE, PT := T#2s); (* Pedestrian crossing grace period *)
            IF Timer.Q THEN
                Timer(IN := FALSE);
                LightState := 1;
            END_IF;
        END_IF;

    1: (* North-South Yellow *)
        NorthSouthYellow := TRUE;
        EastWestRed := TRUE;
        Timer(IN := TRUE, PT := T#2s); (* Yellow light duration *)
        IF Timer.Q THEN
            Timer(IN := FALSE);
            LightState := 2;
        END_IF;

    2: (* East-West Green *)
        EastWestGreen := TRUE;
        NorthSouthRed := TRUE;
        IF PedestrianRequest1 THEN
            PedestrianLight1 := TRUE;
            PedestrianCrossing := NOT (TRUE); (* MUTATED: ASSIGN_NEGATE *)
        END_IF;
        IF PedestrianRequest2 THEN
            PedestrianLight2 := TRUE;
            PedestrianCrossing := TRUE;
        END_IF;
        IF PedestrianCrossing THEN
            Timer(IN := TRUE, PT := T#2s); (* Pedestrian crossing period *)
            IF Timer.Q THEN
                Timer(IN := FALSE);
                PedestrianRequest1 := FALSE;
                PedestrianRequest2 := FALSE;
                PedestrianLight1 := FALSE;
                PedestrianLight2 := FALSE;
                PedestrianCrossing := FALSE;
                LightState := 3;
            END_IF;
        END_IF;

    3: (* East-West Yellow *)
        EastWestYellow := TRUE;
        NorthSouthRed := TRUE;
        Timer(IN := TRUE, PT := T#2s); (* Yellow light duration *)
        IF Timer.Q THEN
            Timer(IN := FALSE);
            LightState := 0;
        END_IF;

END_CASE;

END_FUNCTION_BLOCK

(* ---- M163.st ---- *)
FUNCTION_BLOCK TRAFFIC_CTRL

VAR_INPUT
    PedestrianButton1 : BOOL;
    PedestrianButton2 : BOOL;
END_VAR

VAR_OUTPUT
    NorthSouthRed : BOOL;
    NorthSouthYellow : BOOL;
    NorthSouthGreen : BOOL;
    EastWestRed : BOOL;
    EastWestYellow : BOOL;
    EastWestGreen : BOOL;
    PedestrianLight1 : BOOL;
    PedestrianLight2 : BOOL;
END_VAR

VAR
    LightState : INT := 0; (* 0: North-South Green, 1: North-South Yellow, 2: East-West Green, 3: East-West Yellow *)
    PedestrianRequest1 : BOOL := FALSE;
    PedestrianRequest2 : BOOL := FALSE;
    PedestrianCrossing : BOOL := FALSE;
    Timer : TON;
END_VAR

(* Check for pedestrian requests *)
IF PedestrianButton1 THEN
    PedestrianRequest1 := TRUE;
END_IF;

IF PedestrianButton2 THEN
    PedestrianRequest2 := TRUE;
END_IF;

(* Traffic light state machine *)
CASE LightState OF
    0: (* North-South Green *)
        NorthSouthGreen := TRUE;
        EastWestRed := TRUE;
        IF PedestrianRequest1 OR PedestrianRequest2 THEN
            Timer(IN := TRUE, PT := T#2s); (* Pedestrian crossing grace period *)
            IF Timer.Q THEN
                Timer(IN := FALSE);
                LightState := 1;
            END_IF;
        END_IF;

    1: (* North-South Yellow *)
        NorthSouthYellow := TRUE;
        EastWestRed := TRUE;
        Timer(IN := TRUE, PT := T#2s); (* Yellow light duration *)
        IF Timer.Q THEN
            Timer(IN := FALSE);
            LightState := 2;
        END_IF;

    2: (* East-West Green *)
        EastWestGreen := TRUE;
        NorthSouthRed := TRUE;
        IF PedestrianRequest1 THEN
            PedestrianLight1 := TRUE;
            PedestrianCrossing := TRUE;
        END_IF;
        IF PedestrianRequest2 THEN
            PedestrianLight2 := NOT (TRUE); (* MUTATED: ASSIGN_NEGATE *)
            PedestrianCrossing := TRUE;
        END_IF;
        IF PedestrianCrossing THEN
            Timer(IN := TRUE, PT := T#2s); (* Pedestrian crossing period *)
            IF Timer.Q THEN
                Timer(IN := FALSE);
                PedestrianRequest1 := FALSE;
                PedestrianRequest2 := FALSE;
                PedestrianLight1 := FALSE;
                PedestrianLight2 := FALSE;
                PedestrianCrossing := FALSE;
                LightState := 3;
            END_IF;
        END_IF;

    3: (* East-West Yellow *)
        EastWestYellow := TRUE;
        NorthSouthRed := TRUE;
        Timer(IN := TRUE, PT := T#2s); (* Yellow light duration *)
        IF Timer.Q THEN
            Timer(IN := FALSE);
            LightState := 0;
        END_IF;

END_CASE;

END_FUNCTION_BLOCK

(* ---- M164.st ---- *)
FUNCTION_BLOCK TRAFFIC_CTRL

VAR_INPUT
    PedestrianButton1 : BOOL;
    PedestrianButton2 : BOOL;
END_VAR

VAR_OUTPUT
    NorthSouthRed : BOOL;
    NorthSouthYellow : BOOL;
    NorthSouthGreen : BOOL;
    EastWestRed : BOOL;
    EastWestYellow : BOOL;
    EastWestGreen : BOOL;
    PedestrianLight1 : BOOL;
    PedestrianLight2 : BOOL;
END_VAR

VAR
    LightState : INT := 0; (* 0: North-South Green, 1: North-South Yellow, 2: East-West Green, 3: East-West Yellow *)
    PedestrianRequest1 : BOOL := FALSE;
    PedestrianRequest2 : BOOL := FALSE;
    PedestrianCrossing : BOOL := FALSE;
    Timer : TON;
END_VAR

(* Check for pedestrian requests *)
IF PedestrianButton1 THEN
    PedestrianRequest1 := TRUE;
END_IF;

IF PedestrianButton2 THEN
    PedestrianRequest2 := TRUE;
END_IF;

(* Traffic light state machine *)
CASE LightState OF
    0: (* North-South Green *)
        NorthSouthGreen := TRUE;
        EastWestRed := TRUE;
        IF PedestrianRequest1 OR PedestrianRequest2 THEN
            Timer(IN := TRUE, PT := T#2s); (* Pedestrian crossing grace period *)
            IF Timer.Q THEN
                Timer(IN := FALSE);
                LightState := 1;
            END_IF;
        END_IF;

    1: (* North-South Yellow *)
        NorthSouthYellow := TRUE;
        EastWestRed := TRUE;
        Timer(IN := TRUE, PT := T#2s); (* Yellow light duration *)
        IF Timer.Q THEN
            Timer(IN := FALSE);
            LightState := 2;
        END_IF;

    2: (* East-West Green *)
        EastWestGreen := TRUE;
        NorthSouthRed := TRUE;
        IF PedestrianRequest1 THEN
            PedestrianLight1 := TRUE;
            PedestrianCrossing := TRUE;
        END_IF;
        IF PedestrianRequest2 THEN
            PedestrianLight2 := TRUE;
            PedestrianCrossing := NOT (TRUE); (* MUTATED: ASSIGN_NEGATE *)
        END_IF;
        IF PedestrianCrossing THEN
            Timer(IN := TRUE, PT := T#2s); (* Pedestrian crossing period *)
            IF Timer.Q THEN
                Timer(IN := FALSE);
                PedestrianRequest1 := FALSE;
                PedestrianRequest2 := FALSE;
                PedestrianLight1 := FALSE;
                PedestrianLight2 := FALSE;
                PedestrianCrossing := FALSE;
                LightState := 3;
            END_IF;
        END_IF;

    3: (* East-West Yellow *)
        EastWestYellow := TRUE;
        NorthSouthRed := TRUE;
        Timer(IN := TRUE, PT := T#2s); (* Yellow light duration *)
        IF Timer.Q THEN
            Timer(IN := FALSE);
            LightState := 0;
        END_IF;

END_CASE;

END_FUNCTION_BLOCK

(* ---- M165.st ---- *)
FUNCTION_BLOCK TRAFFIC_CTRL

VAR_INPUT
    PedestrianButton1 : BOOL;
    PedestrianButton2 : BOOL;
END_VAR

VAR_OUTPUT
    NorthSouthRed : BOOL;
    NorthSouthYellow : BOOL;
    NorthSouthGreen : BOOL;
    EastWestRed : BOOL;
    EastWestYellow : BOOL;
    EastWestGreen : BOOL;
    PedestrianLight1 : BOOL;
    PedestrianLight2 : BOOL;
END_VAR

VAR
    LightState : INT := 0; (* 0: North-South Green, 1: North-South Yellow, 2: East-West Green, 3: East-West Yellow *)
    PedestrianRequest1 : BOOL := FALSE;
    PedestrianRequest2 : BOOL := FALSE;
    PedestrianCrossing : BOOL := FALSE;
    Timer : TON;
END_VAR

(* Check for pedestrian requests *)
IF PedestrianButton1 THEN
    PedestrianRequest1 := TRUE;
END_IF;

IF PedestrianButton2 THEN
    PedestrianRequest2 := TRUE;
END_IF;

(* Traffic light state machine *)
CASE LightState OF
    0: (* North-South Green *)
        NorthSouthGreen := TRUE;
        EastWestRed := TRUE;
        IF PedestrianRequest1 OR PedestrianRequest2 THEN
            Timer(IN := TRUE, PT := T#2s); (* Pedestrian crossing grace period *)
            IF Timer.Q THEN
                Timer(IN := FALSE);
                LightState := 1;
            END_IF;
        END_IF;

    1: (* North-South Yellow *)
        NorthSouthYellow := TRUE;
        EastWestRed := TRUE;
        Timer(IN := TRUE, PT := T#2s); (* Yellow light duration *)
        IF Timer.Q THEN
            Timer(IN := FALSE);
            LightState := 2;
        END_IF;

    2: (* East-West Green *)
        EastWestGreen := TRUE;
        NorthSouthRed := TRUE;
        IF PedestrianRequest1 THEN
            PedestrianLight1 := TRUE;
            PedestrianCrossing := TRUE;
        END_IF;
        IF PedestrianRequest2 THEN
            PedestrianLight2 := TRUE;
            PedestrianCrossing := TRUE;
        END_IF;
        IF PedestrianCrossing THEN
            Timer(IN := TRUE, PT := T#2s); (* Pedestrian crossing period *)
            IF Timer.Q THEN
                Timer(IN := FALSE);
                PedestrianRequest1 := NOT (FALSE); (* MUTATED: ASSIGN_NEGATE *)
                PedestrianRequest2 := FALSE;
                PedestrianLight1 := FALSE;
                PedestrianLight2 := FALSE;
                PedestrianCrossing := FALSE;
                LightState := 3;
            END_IF;
        END_IF;

    3: (* East-West Yellow *)
        EastWestYellow := TRUE;
        NorthSouthRed := TRUE;
        Timer(IN := TRUE, PT := T#2s); (* Yellow light duration *)
        IF Timer.Q THEN
            Timer(IN := FALSE);
            LightState := 0;
        END_IF;

END_CASE;

END_FUNCTION_BLOCK

(* ---- M166.st ---- *)
FUNCTION_BLOCK TRAFFIC_CTRL

VAR_INPUT
    PedestrianButton1 : BOOL;
    PedestrianButton2 : BOOL;
END_VAR

VAR_OUTPUT
    NorthSouthRed : BOOL;
    NorthSouthYellow : BOOL;
    NorthSouthGreen : BOOL;
    EastWestRed : BOOL;
    EastWestYellow : BOOL;
    EastWestGreen : BOOL;
    PedestrianLight1 : BOOL;
    PedestrianLight2 : BOOL;
END_VAR

VAR
    LightState : INT := 0; (* 0: North-South Green, 1: North-South Yellow, 2: East-West Green, 3: East-West Yellow *)
    PedestrianRequest1 : BOOL := FALSE;
    PedestrianRequest2 : BOOL := FALSE;
    PedestrianCrossing : BOOL := FALSE;
    Timer : TON;
END_VAR

(* Check for pedestrian requests *)
IF PedestrianButton1 THEN
    PedestrianRequest1 := TRUE;
END_IF;

IF PedestrianButton2 THEN
    PedestrianRequest2 := TRUE;
END_IF;

(* Traffic light state machine *)
CASE LightState OF
    0: (* North-South Green *)
        NorthSouthGreen := TRUE;
        EastWestRed := TRUE;
        IF PedestrianRequest1 OR PedestrianRequest2 THEN
            Timer(IN := TRUE, PT := T#2s); (* Pedestrian crossing grace period *)
            IF Timer.Q THEN
                Timer(IN := FALSE);
                LightState := 1;
            END_IF;
        END_IF;

    1: (* North-South Yellow *)
        NorthSouthYellow := TRUE;
        EastWestRed := TRUE;
        Timer(IN := TRUE, PT := T#2s); (* Yellow light duration *)
        IF Timer.Q THEN
            Timer(IN := FALSE);
            LightState := 2;
        END_IF;

    2: (* East-West Green *)
        EastWestGreen := TRUE;
        NorthSouthRed := TRUE;
        IF PedestrianRequest1 THEN
            PedestrianLight1 := TRUE;
            PedestrianCrossing := TRUE;
        END_IF;
        IF PedestrianRequest2 THEN
            PedestrianLight2 := TRUE;
            PedestrianCrossing := TRUE;
        END_IF;
        IF PedestrianCrossing THEN
            Timer(IN := TRUE, PT := T#2s); (* Pedestrian crossing period *)
            IF Timer.Q THEN
                Timer(IN := FALSE);
                PedestrianRequest1 := FALSE;
                PedestrianRequest2 := NOT (FALSE); (* MUTATED: ASSIGN_NEGATE *)
                PedestrianLight1 := FALSE;
                PedestrianLight2 := FALSE;
                PedestrianCrossing := FALSE;
                LightState := 3;
            END_IF;
        END_IF;

    3: (* East-West Yellow *)
        EastWestYellow := TRUE;
        NorthSouthRed := TRUE;
        Timer(IN := TRUE, PT := T#2s); (* Yellow light duration *)
        IF Timer.Q THEN
            Timer(IN := FALSE);
            LightState := 0;
        END_IF;

END_CASE;

END_FUNCTION_BLOCK

(* ---- M167.st ---- *)
FUNCTION_BLOCK TRAFFIC_CTRL

VAR_INPUT
    PedestrianButton1 : BOOL;
    PedestrianButton2 : BOOL;
END_VAR

VAR_OUTPUT
    NorthSouthRed : BOOL;
    NorthSouthYellow : BOOL;
    NorthSouthGreen : BOOL;
    EastWestRed : BOOL;
    EastWestYellow : BOOL;
    EastWestGreen : BOOL;
    PedestrianLight1 : BOOL;
    PedestrianLight2 : BOOL;
END_VAR

VAR
    LightState : INT := 0; (* 0: North-South Green, 1: North-South Yellow, 2: East-West Green, 3: East-West Yellow *)
    PedestrianRequest1 : BOOL := FALSE;
    PedestrianRequest2 : BOOL := FALSE;
    PedestrianCrossing : BOOL := FALSE;
    Timer : TON;
END_VAR

(* Check for pedestrian requests *)
IF PedestrianButton1 THEN
    PedestrianRequest1 := TRUE;
END_IF;

IF PedestrianButton2 THEN
    PedestrianRequest2 := TRUE;
END_IF;

(* Traffic light state machine *)
CASE LightState OF
    0: (* North-South Green *)
        NorthSouthGreen := TRUE;
        EastWestRed := TRUE;
        IF PedestrianRequest1 OR PedestrianRequest2 THEN
            Timer(IN := TRUE, PT := T#2s); (* Pedestrian crossing grace period *)
            IF Timer.Q THEN
                Timer(IN := FALSE);
                LightState := 1;
            END_IF;
        END_IF;

    1: (* North-South Yellow *)
        NorthSouthYellow := TRUE;
        EastWestRed := TRUE;
        Timer(IN := TRUE, PT := T#2s); (* Yellow light duration *)
        IF Timer.Q THEN
            Timer(IN := FALSE);
            LightState := 2;
        END_IF;

    2: (* East-West Green *)
        EastWestGreen := TRUE;
        NorthSouthRed := TRUE;
        IF PedestrianRequest1 THEN
            PedestrianLight1 := TRUE;
            PedestrianCrossing := TRUE;
        END_IF;
        IF PedestrianRequest2 THEN
            PedestrianLight2 := TRUE;
            PedestrianCrossing := TRUE;
        END_IF;
        IF PedestrianCrossing THEN
            Timer(IN := TRUE, PT := T#2s); (* Pedestrian crossing period *)
            IF Timer.Q THEN
                Timer(IN := FALSE);
                PedestrianRequest1 := FALSE;
                PedestrianRequest2 := FALSE;
                PedestrianLight1 := NOT (FALSE); (* MUTATED: ASSIGN_NEGATE *)
                PedestrianLight2 := FALSE;
                PedestrianCrossing := FALSE;
                LightState := 3;
            END_IF;
        END_IF;

    3: (* East-West Yellow *)
        EastWestYellow := TRUE;
        NorthSouthRed := TRUE;
        Timer(IN := TRUE, PT := T#2s); (* Yellow light duration *)
        IF Timer.Q THEN
            Timer(IN := FALSE);
            LightState := 0;
        END_IF;

END_CASE;

END_FUNCTION_BLOCK

(* ---- M168.st ---- *)
FUNCTION_BLOCK TRAFFIC_CTRL

VAR_INPUT
    PedestrianButton1 : BOOL;
    PedestrianButton2 : BOOL;
END_VAR

VAR_OUTPUT
    NorthSouthRed : BOOL;
    NorthSouthYellow : BOOL;
    NorthSouthGreen : BOOL;
    EastWestRed : BOOL;
    EastWestYellow : BOOL;
    EastWestGreen : BOOL;
    PedestrianLight1 : BOOL;
    PedestrianLight2 : BOOL;
END_VAR

VAR
    LightState : INT := 0; (* 0: North-South Green, 1: North-South Yellow, 2: East-West Green, 3: East-West Yellow *)
    PedestrianRequest1 : BOOL := FALSE;
    PedestrianRequest2 : BOOL := FALSE;
    PedestrianCrossing : BOOL := FALSE;
    Timer : TON;
END_VAR

(* Check for pedestrian requests *)
IF PedestrianButton1 THEN
    PedestrianRequest1 := TRUE;
END_IF;

IF PedestrianButton2 THEN
    PedestrianRequest2 := TRUE;
END_IF;

(* Traffic light state machine *)
CASE LightState OF
    0: (* North-South Green *)
        NorthSouthGreen := TRUE;
        EastWestRed := TRUE;
        IF PedestrianRequest1 OR PedestrianRequest2 THEN
            Timer(IN := TRUE, PT := T#2s); (* Pedestrian crossing grace period *)
            IF Timer.Q THEN
                Timer(IN := FALSE);
                LightState := 1;
            END_IF;
        END_IF;

    1: (* North-South Yellow *)
        NorthSouthYellow := TRUE;
        EastWestRed := TRUE;
        Timer(IN := TRUE, PT := T#2s); (* Yellow light duration *)
        IF Timer.Q THEN
            Timer(IN := FALSE);
            LightState := 2;
        END_IF;

    2: (* East-West Green *)
        EastWestGreen := TRUE;
        NorthSouthRed := TRUE;
        IF PedestrianRequest1 THEN
            PedestrianLight1 := TRUE;
            PedestrianCrossing := TRUE;
        END_IF;
        IF PedestrianRequest2 THEN
            PedestrianLight2 := TRUE;
            PedestrianCrossing := TRUE;
        END_IF;
        IF PedestrianCrossing THEN
            Timer(IN := TRUE, PT := T#2s); (* Pedestrian crossing period *)
            IF Timer.Q THEN
                Timer(IN := FALSE);
                PedestrianRequest1 := FALSE;
                PedestrianRequest2 := FALSE;
                PedestrianLight1 := FALSE;
                PedestrianLight2 := NOT (FALSE); (* MUTATED: ASSIGN_NEGATE *)
                PedestrianCrossing := FALSE;
                LightState := 3;
            END_IF;
        END_IF;

    3: (* East-West Yellow *)
        EastWestYellow := TRUE;
        NorthSouthRed := TRUE;
        Timer(IN := TRUE, PT := T#2s); (* Yellow light duration *)
        IF Timer.Q THEN
            Timer(IN := FALSE);
            LightState := 0;
        END_IF;

END_CASE;

END_FUNCTION_BLOCK
